REGION Network 17: Sinais Main Line POSTO 80
   // JOB [0]=- ANDON;
   // JOB [1] = EMERGÊNCIA;
   // JOB [2] = AP SUP FREIO;
   // JOB [3] = PY EXCENTRIO;
   // JOB [4] = PY CUBO DISCO
   RUNG wire#powerrail
      Contact( "Get Sinais de Interlock Main line".Station[1]."Sinal do job"[0] )
      I_Contact( "BYPASS_MOD_2" )
      I_Contact( "BYPASS_GERAL" )
      I_Contact( "BYPASS_POSTO_80" )
      Coil( "Signals".ProcessInterlock_APLC_Input[1].ModezoneInterlock_APLC_Input[2].StationInterlock_APLC_Input[3].PositionInterlock_APLC_Input[1].EquipmentInterlock_APLC_Input[1].SignalInterlock_APLC_Input[1] )
   END_RUNG
   RUNG wire#powerrail
      Contact( "Get Sinais de Interlock Main line".Station[1]."Sinal do job"[1] )
      I_Contact( "BYPASS_MOD_2" )
      I_Contact( "BYPASS_GERAL" )
      I_Contact( "BYPASS_POSTO_80" )
      Coil( "Signals".ProcessInterlock_APLC_Input[1].ModezoneInterlock_APLC_Input[2].StationInterlock_APLC_Input[3].PositionInterlock_APLC_Input[1].EquipmentInterlock_APLC_Input[1].SignalInterlock_APLC_Input[2] )
   END_RUNG
   // the same network as SCL:
   "Signals".ProcessInterlock_APLC_Input[1].ModezoneInterlock_APLC_Input[2].StationInterlock_APLC_Input[3].PositionInterlock_APLC_Input[1].EquipmentInterlock_APLC_Input[1].SignalInterlock_APLC_Input[1] := "Get Sinais de Interlock Main line".Station[1]."Sinal do job"[0] AND NOT "BYPASS_MOD_2" AND NOT "BYPASS_GERAL" AND NOT "BYPASS_POSTO_80";
   "Signals".ProcessInterlock_APLC_Input[1].ModezoneInterlock_APLC_Input[2].StationInterlock_APLC_Input[3].PositionInterlock_APLC_Input[1].EquipmentInterlock_APLC_Input[1].SignalInterlock_APLC_Input[2] := "Get Sinais de Interlock Main line".Station[1]."Sinal do job"[1] AND NOT "BYPASS_MOD_2" AND NOT "BYPASS_GERAL" AND NOT "BYPASS_POSTO_80";
END_REGION

REGION Network 18: Sinais Main Line POSTO 90
   // JOB [0] = ANDON;
   // JOB [1] = EMERGÊNCIA;
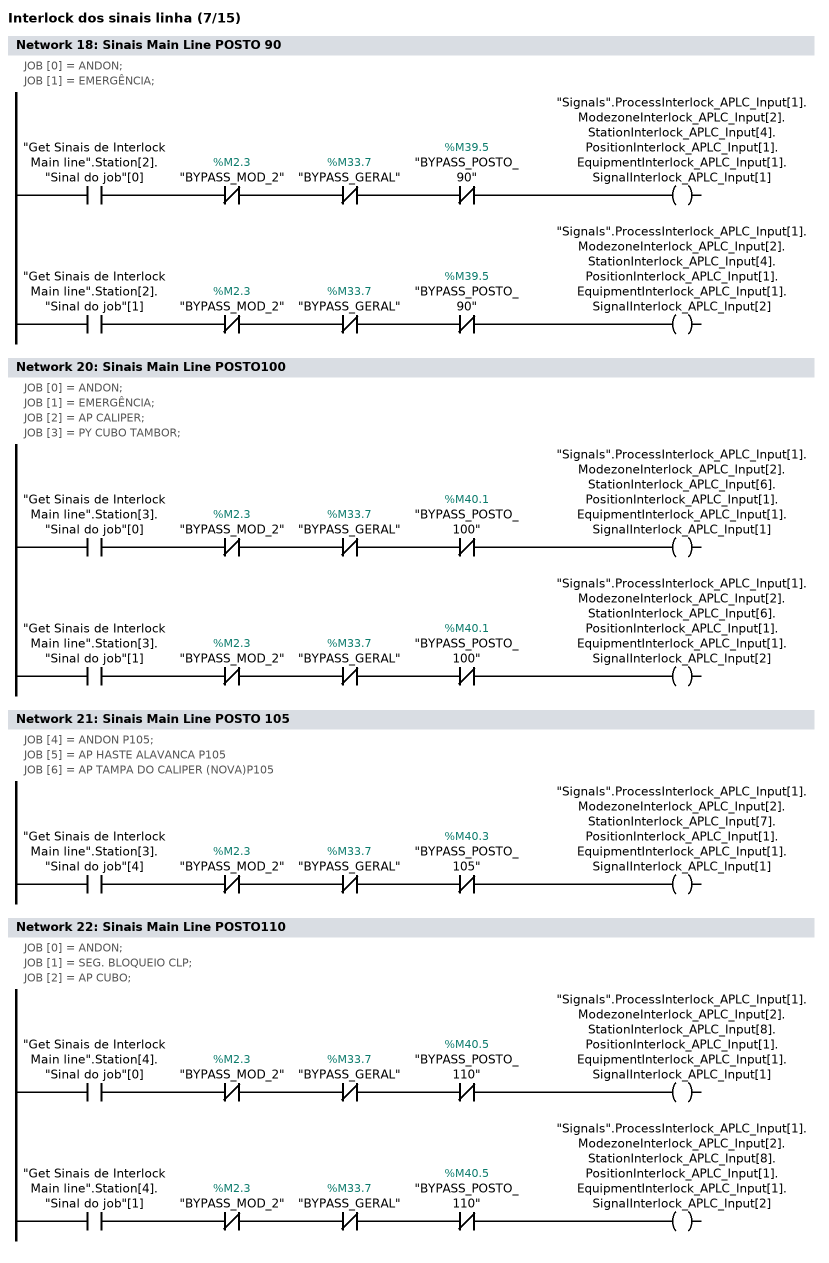
   RUNG wire#powerrail
      Contact( "Get Sinais de Interlock Main line".Station[2]."Sinal do job"[0] )
      I_Contact( "BYPASS_MOD_2" )
      I_Contact( "BYPASS_GERAL" )
      I_Contact( "BYPASS_POSTO_90" )
      Coil( "Signals".ProcessInterlock_APLC_Input[1].ModezoneInterlock_APLC_Input[2].StationInterlock_APLC_Input[4].PositionInterlock_APLC_Input[1].EquipmentInterlock_APLC_Input[1].SignalInterlock_APLC_Input[1] )
   END_RUNG
   RUNG wire#powerrail
      Contact( "Get Sinais de Interlock Main line".Station[2]."Sinal do job"[1] )
      I_Contact( "BYPASS_MOD_2" )
      I_Contact( "BYPASS_GERAL" )
      I_Contact( "BYPASS_POSTO_90" )
      Coil( "Signals".ProcessInterlock_APLC_Input[1].ModezoneInterlock_APLC_Input[2].StationInterlock_APLC_Input[4].PositionInterlock_APLC_Input[1].EquipmentInterlock_APLC_Input[1].SignalInterlock_APLC_Input[2] )
   END_RUNG
   // the same network as SCL:
   "Signals".ProcessInterlock_APLC_Input[1].ModezoneInterlock_APLC_Input[2].StationInterlock_APLC_Input[4].PositionInterlock_APLC_Input[1].EquipmentInterlock_APLC_Input[1].SignalInterlock_APLC_Input[1] := "Get Sinais de Interlock Main line".Station[2]."Sinal do job"[0] AND NOT "BYPASS_MOD_2" AND NOT "BYPASS_GERAL" AND NOT "BYPASS_POSTO_90";
   "Signals".ProcessInterlock_APLC_Input[1].ModezoneInterlock_APLC_Input[2].StationInterlock_APLC_Input[4].PositionInterlock_APLC_Input[1].EquipmentInterlock_APLC_Input[1].SignalInterlock_APLC_Input[2] := "Get Sinais de Interlock Main line".Station[2]."Sinal do job"[1] AND NOT "BYPASS_MOD_2" AND NOT "BYPASS_GERAL" AND NOT "BYPASS_POSTO_90";
END_REGION

REGION Network 19: Sinais Main Line POSTO 95
   // JOB [2] = AP HOLDER. P95
END_REGION

REGION Network 20: Sinais Main Line POSTO100
   // JOB [0] = ANDON;
   // JOB [1] = EMERGÊNCIA;
   // JOB [2] = AP CALIPER;
   // JOB [3] = PY CUBO TAMBOR;
   RUNG wire#powerrail
      Contact( "Get Sinais de Interlock Main line".Station[3]."Sinal do job"[0] )
      I_Contact( "BYPASS_MOD_2" )
      I_Contact( "BYPASS_GERAL" )
      I_Contact( "BYPASS_POSTO_100" )
      Coil( "Signals".ProcessInterlock_APLC_Input[1].ModezoneInterlock_APLC_Input[2].StationInterlock_APLC_Input[6].PositionInterlock_APLC_Input[1].EquipmentInterlock_APLC_Input[1].SignalInterlock_APLC_Input[1] )
   END_RUNG
   RUNG wire#powerrail
      Contact( "Get Sinais de Interlock Main line".Station[3]."Sinal do job"[1] )
      I_Contact( "BYPASS_MOD_2" )
      I_Contact( "BYPASS_GERAL" )
      I_Contact( "BYPASS_POSTO_100" )
      Coil( "Signals".ProcessInterlock_APLC_Input[1].ModezoneInterlock_APLC_Input[2].StationInterlock_APLC_Input[6].PositionInterlock_APLC_Input[1].EquipmentInterlock_APLC_Input[1].SignalInterlock_APLC_Input[2] )
   END_RUNG
   // the same network as SCL:
   "Signals".ProcessInterlock_APLC_Input[1].ModezoneInterlock_APLC_Input[2].StationInterlock_APLC_Input[6].PositionInterlock_APLC_Input[1].EquipmentInterlock_APLC_Input[1].SignalInterlock_APLC_Input[1] := "Get Sinais de Interlock Main line".Station[3]."Sinal do job"[0] AND NOT "BYPASS_MOD_2" AND NOT "BYPASS_GERAL" AND NOT "BYPASS_POSTO_100";
   "Signals".ProcessInterlock_APLC_Input[1].ModezoneInterlock_APLC_Input[2].StationInterlock_APLC_Input[6].PositionInterlock_APLC_Input[1].EquipmentInterlock_APLC_Input[1].SignalInterlock_APLC_Input[2] := "Get Sinais de Interlock Main line".Station[3]."Sinal do job"[1] AND NOT "BYPASS_MOD_2" AND NOT "BYPASS_GERAL" AND NOT "BYPASS_POSTO_100";
END_REGION

REGION Network 21: Sinais Main Line POSTO 105
   // JOB [4] = ANDON P105;
   // JOB [5] = AP HASTE ALAVANCA P105
   // JOB [6] = AP TAMPA DO CALIPER (NOVA)P105
   RUNG wire#powerrail
      Contact( "Get Sinais de Interlock Main line".Station[3]."Sinal do job"[4] )
      I_Contact( "BYPASS_MOD_2" )
      I_Contact( "BYPASS_GERAL" )
      I_Contact( "BYPASS_POSTO_105" )
      Coil( "Signals".ProcessInterlock_APLC_Input[1].ModezoneInterlock_APLC_Input[2].StationInterlock_APLC_Input[7].PositionInterlock_APLC_Input[1].EquipmentInterlock_APLC_Input[1].SignalInterlock_APLC_Input[1] )
   END_RUNG
   // the same network as SCL:
   "Signals".ProcessInterlock_APLC_Input[1].ModezoneInterlock_APLC_Input[2].StationInterlock_APLC_Input[7].PositionInterlock_APLC_Input[1].EquipmentInterlock_APLC_Input[1].SignalInterlock_APLC_Input[1] := "Get Sinais de Interlock Main line".Station[3]."Sinal do job"[4] AND NOT "BYPASS_MOD_2" AND NOT "BYPASS_GERAL" AND NOT "BYPASS_POSTO_105";
END_REGION

REGION Network 22: Sinais Main Line POSTO110
   // JOB [0] = ANDON;
   // JOB [1] = SEG. BLOQUEIO CLP;
   // JOB [2] = AP CUBO;
   RUNG wire#powerrail
      Contact( "Get Sinais de Interlock Main line".Station[4]."Sinal do job"[0] )
      I_Contact( "BYPASS_MOD_2" )
      I_Contact( "BYPASS_GERAL" )
      I_Contact( "BYPASS_POSTO_110" )
      Coil( "Signals".ProcessInterlock_APLC_Input[1].ModezoneInterlock_APLC_Input[2].StationInterlock_APLC_Input[8].PositionInterlock_APLC_Input[1].EquipmentInterlock_APLC_Input[1].SignalInterlock_APLC_Input[1] )
   END_RUNG
   RUNG wire#powerrail
      Contact( "Get Sinais de Interlock Main line".Station[4]."Sinal do job"[1] )
      I_Contact( "BYPASS_MOD_2" )
      I_Contact( "BYPASS_GERAL" )
      I_Contact( "BYPASS_POSTO_110" )
      Coil( "Signals".ProcessInterlock_APLC_Input[1].ModezoneInterlock_APLC_Input[2].StationInterlock_APLC_Input[8].PositionInterlock_APLC_Input[1].EquipmentInterlock_APLC_Input[1].SignalInterlock_APLC_Input[2] )
   END_RUNG
   // the same network as SCL:
   "Signals".ProcessInterlock_APLC_Input[1].ModezoneInterlock_APLC_Input[2].StationInterlock_APLC_Input[8].PositionInterlock_APLC_Input[1].EquipmentInterlock_APLC_Input[1].SignalInterlock_APLC_Input[1] := "Get Sinais de Interlock Main line".Station[4]."Sinal do job"[0] AND NOT "BYPASS_MOD_2" AND NOT "BYPASS_GERAL" AND NOT "BYPASS_POSTO_110";
   "Signals".ProcessInterlock_APLC_Input[1].ModezoneInterlock_APLC_Input[2].StationInterlock_APLC_Input[8].PositionInterlock_APLC_Input[1].EquipmentInterlock_APLC_Input[1].SignalInterlock_APLC_Input[2] := "Get Sinais de Interlock Main line".Station[4]."Sinal do job"[1] AND NOT "BYPASS_MOD_2" AND NOT "BYPASS_GERAL" AND NOT "BYPASS_POSTO_110";
END_REGION

REGION Network 23: Sinais Main Line POSTO 115
   // JOB [3] = ANDON P115;
   // JOB [4] = CRAVADOR.
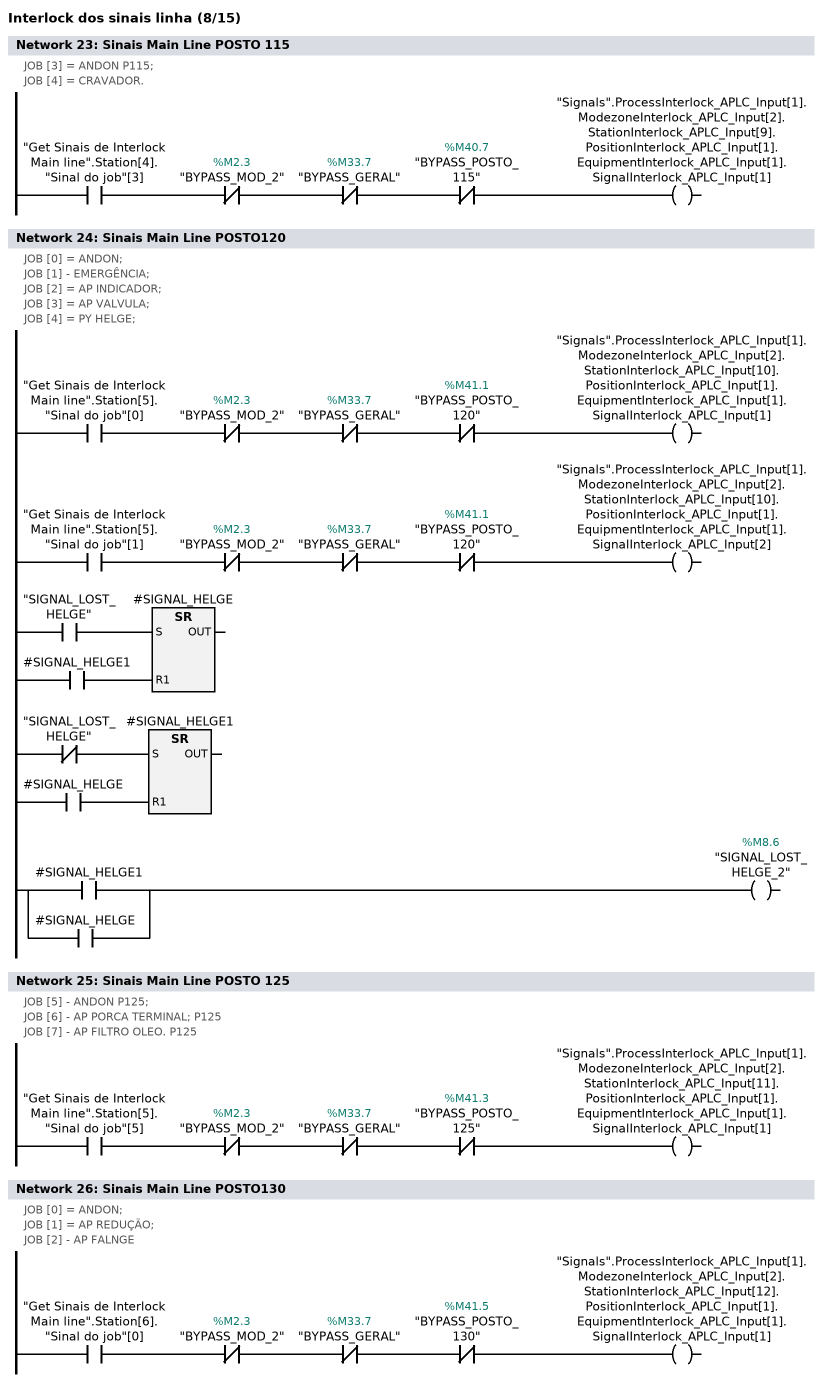
   RUNG wire#powerrail
      Contact( "Get Sinais de Interlock Main line".Station[4]."Sinal do job"[3] )
      I_Contact( "BYPASS_MOD_2" )
      I_Contact( "BYPASS_GERAL" )
      I_Contact( "BYPASS_POSTO_115" )
      Coil( "Signals".ProcessInterlock_APLC_Input[1].ModezoneInterlock_APLC_Input[2].StationInterlock_APLC_Input[9].PositionInterlock_APLC_Input[1].EquipmentInterlock_APLC_Input[1].SignalInterlock_APLC_Input[1] )
   END_RUNG
   // the same network as SCL:
   "Signals".ProcessInterlock_APLC_Input[1].ModezoneInterlock_APLC_Input[2].StationInterlock_APLC_Input[9].PositionInterlock_APLC_Input[1].EquipmentInterlock_APLC_Input[1].SignalInterlock_APLC_Input[1] := "Get Sinais de Interlock Main line".Station[4]."Sinal do job"[3] AND NOT "BYPASS_MOD_2" AND NOT "BYPASS_GERAL" AND NOT "BYPASS_POSTO_115";
END_REGION

REGION Network 24: Sinais Main Line POSTO120
   // JOB [0] = ANDON;
   // JOB [1] - EMERGÊNCIA;
   // JOB [2] = AP INDICADOR;
   // JOB [3] = AP VALVULA;
   // JOB [4] = PY HELGE;
   RUNG wire#powerrail
      Contact( "Get Sinais de Interlock Main line".Station[5]."Sinal do job"[0] )
      I_Contact( "BYPASS_MOD_2" )
      I_Contact( "BYPASS_GERAL" )
      I_Contact( "BYPASS_POSTO_120" )
      Coil( "Signals".ProcessInterlock_APLC_Input[1].ModezoneInterlock_APLC_Input[2].StationInterlock_APLC_Input[10].PositionInterlock_APLC_Input[1].EquipmentInterlock_APLC_Input[1].SignalInterlock_APLC_Input[1] )
   END_RUNG
   RUNG wire#powerrail
      Contact( "Get Sinais de Interlock Main line".Station[5]."Sinal do job"[1] )
      I_Contact( "BYPASS_MOD_2" )
      I_Contact( "BYPASS_GERAL" )
      I_Contact( "BYPASS_POSTO_120" )
      Coil( "Signals".ProcessInterlock_APLC_Input[1].ModezoneInterlock_APLC_Input[2].StationInterlock_APLC_Input[10].PositionInterlock_APLC_Input[1].EquipmentInterlock_APLC_Input[1].SignalInterlock_APLC_Input[2] )
   END_RUNG
   RUNG wire#powerrail
      Contact( "SIGNAL_LOST_HELGE" )
      S_SR(operand := #SIGNAL_HELGE, r1 := wire#w1)
   END_RUNG
   RUNG wire#powerrail
      Contact( #SIGNAL_HELGE1 )
   END_RUNG wire#w1
   RUNG wire#powerrail
      I_Contact( "SIGNAL_LOST_HELGE" )
      S_SR(operand := #SIGNAL_HELGE1, r1 := wire#w2)
   END_RUNG
   RUNG wire#powerrail
      Contact( #SIGNAL_HELGE )
   END_RUNG wire#w2
   RUNG wire#powerrail
      Contact( #SIGNAL_HELGE1 )
      wire#w3
      Coil( "SIGNAL_LOST_HELGE_2" )
   END_RUNG
   RUNG wire#powerrail
      Contact( #SIGNAL_HELGE )
   END_RUNG wire#w3
   // the same network as SCL:
   "Signals".ProcessInterlock_APLC_Input[1].ModezoneInterlock_APLC_Input[2].StationInterlock_APLC_Input[10].PositionInterlock_APLC_Input[1].EquipmentInterlock_APLC_Input[1].SignalInterlock_APLC_Input[1] := "Get Sinais de Interlock Main line".Station[5]."Sinal do job"[0] AND NOT "BYPASS_MOD_2" AND NOT "BYPASS_GERAL" AND NOT "BYPASS_POSTO_120";
   "Signals".ProcessInterlock_APLC_Input[1].ModezoneInterlock_APLC_Input[2].StationInterlock_APLC_Input[10].PositionInterlock_APLC_Input[1].EquipmentInterlock_APLC_Input[1].SignalInterlock_APLC_Input[2] := "Get Sinais de Interlock Main line".Station[5]."Sinal do job"[1] AND NOT "BYPASS_MOD_2" AND NOT "BYPASS_GERAL" AND NOT "BYPASS_POSTO_120";
   IF "SIGNAL_LOST_HELGE" THEN
       #SIGNAL_HELGE := TRUE;   // SR flip-flop
   END_IF;
   IF #SIGNAL_HELGE1 THEN #SIGNAL_HELGE := FALSE; END_IF;
   IF NOT "SIGNAL_LOST_HELGE" THEN
       #SIGNAL_HELGE1 := TRUE;   // SR flip-flop
   END_IF;
   IF #SIGNAL_HELGE THEN #SIGNAL_HELGE1 := FALSE; END_IF;
   "SIGNAL_LOST_HELGE_2" := #SIGNAL_HELGE1 OR #SIGNAL_HELGE;
END_REGION

REGION Network 25: Sinais Main Line POSTO 125
   // JOB [5] - ANDON P125;
   // JOB [6] - AP PORCA TERMINAL; P125
   // JOB [7] - AP FILTRO OLEO. P125
   RUNG wire#powerrail
      Contact( "Get Sinais de Interlock Main line".Station[5]."Sinal do job"[5] )
      I_Contact( "BYPASS_MOD_2" )
      I_Contact( "BYPASS_GERAL" )
      I_Contact( "BYPASS_POSTO_125" )
      Coil( "Signals".ProcessInterlock_APLC_Input[1].ModezoneInterlock_APLC_Input[2].StationInterlock_APLC_Input[11].PositionInterlock_APLC_Input[1].EquipmentInterlock_APLC_Input[1].SignalInterlock_APLC_Input[1] )
   END_RUNG
   // the same network as SCL:
   "Signals".ProcessInterlock_APLC_Input[1].ModezoneInterlock_APLC_Input[2].StationInterlock_APLC_Input[11].PositionInterlock_APLC_Input[1].EquipmentInterlock_APLC_Input[1].SignalInterlock_APLC_Input[1] := "Get Sinais de Interlock Main line".Station[5]."Sinal do job"[5] AND NOT "BYPASS_MOD_2" AND NOT "BYPASS_GERAL" AND NOT "BYPASS_POSTO_125";
END_REGION

REGION Network 26: Sinais Main Line POSTO130
   // JOB [0] = ANDON;
   // JOB [1] = AP REDUÇÃO;
   // JOB [2] - AP FALNGE
   RUNG wire#powerrail
      Contact( "Get Sinais de Interlock Main line".Station[6]."Sinal do job"[0] )
      I_Contact( "BYPASS_MOD_2" )
      I_Contact( "BYPASS_GERAL" )
      I_Contact( "BYPASS_POSTO_130" )
      Coil( "Signals".ProcessInterlock_APLC_Input[1].ModezoneInterlock_APLC_Input[2].StationInterlock_APLC_Input[12].PositionInterlock_APLC_Input[1].EquipmentInterlock_APLC_Input[1].SignalInterlock_APLC_Input[1] )
   END_RUNG
   // the same network as SCL:
   "Signals".ProcessInterlock_APLC_Input[1].ModezoneInterlock_APLC_Input[2].StationInterlock_APLC_Input[12].PositionInterlock_APLC_Input[1].EquipmentInterlock_APLC_Input[1].SignalInterlock_APLC_Input[1] := "Get Sinais de Interlock Main line".Station[6]."Sinal do job"[0] AND NOT "BYPASS_MOD_2" AND NOT "BYPASS_GERAL" AND NOT "BYPASS_POSTO_130";
END_REGION

REGION Network 27: Sinais Main Line POSTO140
   // JOB [0] = ANDON;
   // JOB [1] = EMERGÊNCIA;
   // JOB [2] = ESTANQUEIDADE CILINDRO;
   // JOB [3] = ESTANQUEIDADE CARCAÇA.
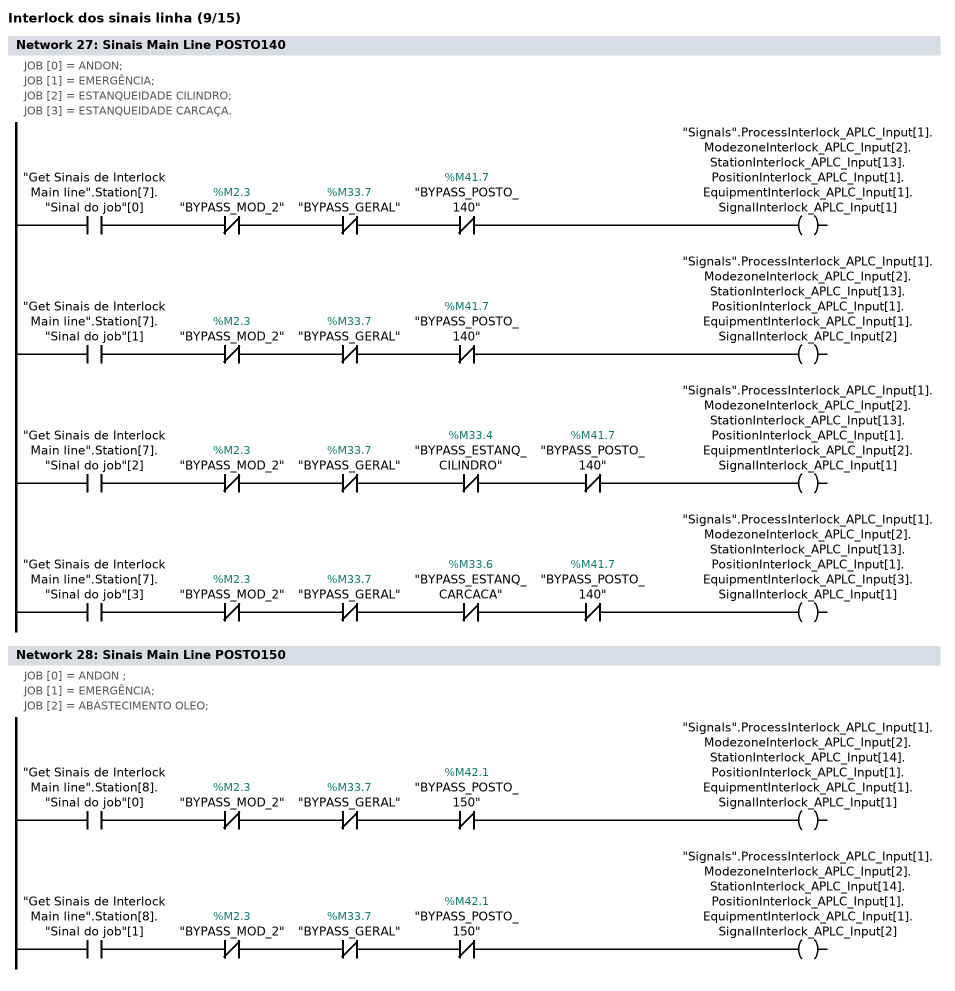
   RUNG wire#powerrail
      Contact( "Get Sinais de Interlock Main line".Station[7]."Sinal do job"[0] )
      I_Contact( "BYPASS_MOD_2" )
      I_Contact( "BYPASS_GERAL" )
      I_Contact( "BYPASS_POSTO_140" )
      Coil( "Signals".ProcessInterlock_APLC_Input[1].ModezoneInterlock_APLC_Input[2].StationInterlock_APLC_Input[13].PositionInterlock_APLC_Input[1].EquipmentInterlock_APLC_Input[1].SignalInterlock_APLC_Input[1] )
   END_RUNG
   RUNG wire#powerrail
      Contact( "Get Sinais de Interlock Main line".Station[7]."Sinal do job"[1] )
      I_Contact( "BYPASS_MOD_2" )
      I_Contact( "BYPASS_GERAL" )
      I_Contact( "BYPASS_POSTO_140" )
      Coil( "Signals".ProcessInterlock_APLC_Input[1].ModezoneInterlock_APLC_Input[2].StationInterlock_APLC_Input[13].PositionInterlock_APLC_Input[1].EquipmentInterlock_APLC_Input[1].SignalInterlock_APLC_Input[2] )
   END_RUNG
   RUNG wire#powerrail
      Contact( "Get Sinais de Interlock Main line".Station[7]."Sinal do job"[2] )
      I_Contact( "BYPASS_MOD_2" )
      I_Contact( "BYPASS_GERAL" )
      I_Contact( "BYPASS_ESTANQ_CILINDRO" )
      I_Contact( "BYPASS_POSTO_140" )
      Coil( "Signals".ProcessInterlock_APLC_Input[1].ModezoneInterlock_APLC_Input[2].StationInterlock_APLC_Input[13].PositionInterlock_APLC_Input[1].EquipmentInterlock_APLC_Input[2].SignalInterlock_APLC_Input[1] )
   END_RUNG
   RUNG wire#powerrail
      Contact( "Get Sinais de Interlock Main line".Station[7]."Sinal do job"[3] )
      I_Contact( "BYPASS_MOD_2" )
      I_Contact( "BYPASS_GERAL" )
      I_Contact( "BYPASS_ESTANQ_CARCACA" )
      I_Contact( "BYPASS_POSTO_140" )
      Coil( "Signals".ProcessInterlock_APLC_Input[1].ModezoneInterlock_APLC_Input[2].StationInterlock_APLC_Input[13].PositionInterlock_APLC_Input[1].EquipmentInterlock_APLC_Input[3].SignalInterlock_APLC_Input[1] )
   END_RUNG
   // the same network as SCL:
   "Signals".ProcessInterlock_APLC_Input[1].ModezoneInterlock_APLC_Input[2].StationInterlock_APLC_Input[13].PositionInterlock_APLC_Input[1].EquipmentInterlock_APLC_Input[1].SignalInterlock_APLC_Input[1] := "Get Sinais de Interlock Main line".Station[7]."Sinal do job"[0] AND NOT "BYPASS_MOD_2" AND NOT "BYPASS_GERAL" AND NOT "BYPASS_POSTO_140";
   "Signals".ProcessInterlock_APLC_Input[1].ModezoneInterlock_APLC_Input[2].StationInterlock_APLC_Input[13].PositionInterlock_APLC_Input[1].EquipmentInterlock_APLC_Input[1].SignalInterlock_APLC_Input[2] := "Get Sinais de Interlock Main line".Station[7]."Sinal do job"[1] AND NOT "BYPASS_MOD_2" AND NOT "BYPASS_GERAL" AND NOT "BYPASS_POSTO_140";
   "Signals".ProcessInterlock_APLC_Input[1].ModezoneInterlock_APLC_Input[2].StationInterlock_APLC_Input[13].PositionInterlock_APLC_Input[1].EquipmentInterlock_APLC_Input[2].SignalInterlock_APLC_Input[1] := "Get Sinais de Interlock Main line".Station[7]."Sinal do job"[2] AND NOT "BYPASS_MOD_2" AND NOT "BYPASS_GERAL" AND NOT "BYPASS_ESTANQ_CILINDRO" AND NOT "BYPASS_POSTO_140";
   "Signals".ProcessInterlock_APLC_Input[1].ModezoneInterlock_APLC_Input[2].StationInterlock_APLC_Input[13].PositionInterlock_APLC_Input[1].EquipmentInterlock_APLC_Input[3].SignalInterlock_APLC_Input[1] := "Get Sinais de Interlock Main line".Station[7]."Sinal do job"[3] AND NOT "BYPASS_MOD_2" AND NOT "BYPASS_GERAL" AND NOT "BYPASS_ESTANQ_CARCACA" AND NOT "BYPASS_POSTO_140";
END_REGION

REGION Network 28: Sinais Main Line POSTO150
   // JOB [0] = ANDON ;
   // JOB [1] = EMERGÊNCIA;
   // JOB [2] = ABASTECIMENTO OLEO;
   RUNG wire#powerrail
      Contact( "Get Sinais de Interlock Main line".Station[8]."Sinal do job"[0] )
      I_Contact( "BYPASS_MOD_2" )
      I_Contact( "BYPASS_GERAL" )
      I_Contact( "BYPASS_POSTO_150" )
      Coil( "Signals".ProcessInterlock_APLC_Input[1].ModezoneInterlock_APLC_Input[2].StationInterlock_APLC_Input[14].PositionInterlock_APLC_Input[1].EquipmentInterlock_APLC_Input[1].SignalInterlock_APLC_Input[1] )
   END_RUNG
   RUNG wire#powerrail
      Contact( "Get Sinais de Interlock Main line".Station[8]."Sinal do job"[1] )
      I_Contact( "BYPASS_MOD_2" )
      I_Contact( "BYPASS_GERAL" )
      I_Contact( "BYPASS_POSTO_150" )
      Coil( "Signals".ProcessInterlock_APLC_Input[1].ModezoneInterlock_APLC_Input[2].StationInterlock_APLC_Input[14].PositionInterlock_APLC_Input[1].EquipmentInterlock_APLC_Input[1].SignalInterlock_APLC_Input[2] )
   END_RUNG
   // the same network as SCL:
   "Signals".ProcessInterlock_APLC_Input[1].ModezoneInterlock_APLC_Input[2].StationInterlock_APLC_Input[14].PositionInterlock_APLC_Input[1].EquipmentInterlock_APLC_Input[1].SignalInterlock_APLC_Input[1] := "Get Sinais de Interlock Main line".Station[8]."Sinal do job"[0] AND NOT "BYPASS_MOD_2" AND NOT "BYPASS_GERAL" AND NOT "BYPASS_POSTO_150";
   "Signals".ProcessInterlock_APLC_Input[1].ModezoneInterlock_APLC_Input[2].StationInterlock_APLC_Input[14].PositionInterlock_APLC_Input[1].EquipmentInterlock_APLC_Input[1].SignalInterlock_APLC_Input[2] := "Get Sinais de Interlock Main line".Station[8]."Sinal do job"[1] AND NOT "BYPASS_MOD_2" AND NOT "BYPASS_GERAL" AND NOT "BYPASS_POSTO_150";
END_REGION

REGION Network 29: Sinais Main Line Q.G
   // JOB [0] = ANDON;
   // JOB [1] = EMERGÊNCIA;
   // JOB [2] - EIXO PENDURADO;
   // JOB [3] - GAP PRESENTE CAB;
   // JOB [4] - GAP PRESENTE TAKT 
   // STATION 10 JOB [0] = TRANSPORTADOR EM MANUAL
   // GAP + EIXO PENDURADO
   // MODEZONE 1 PARADO (FALCARE)
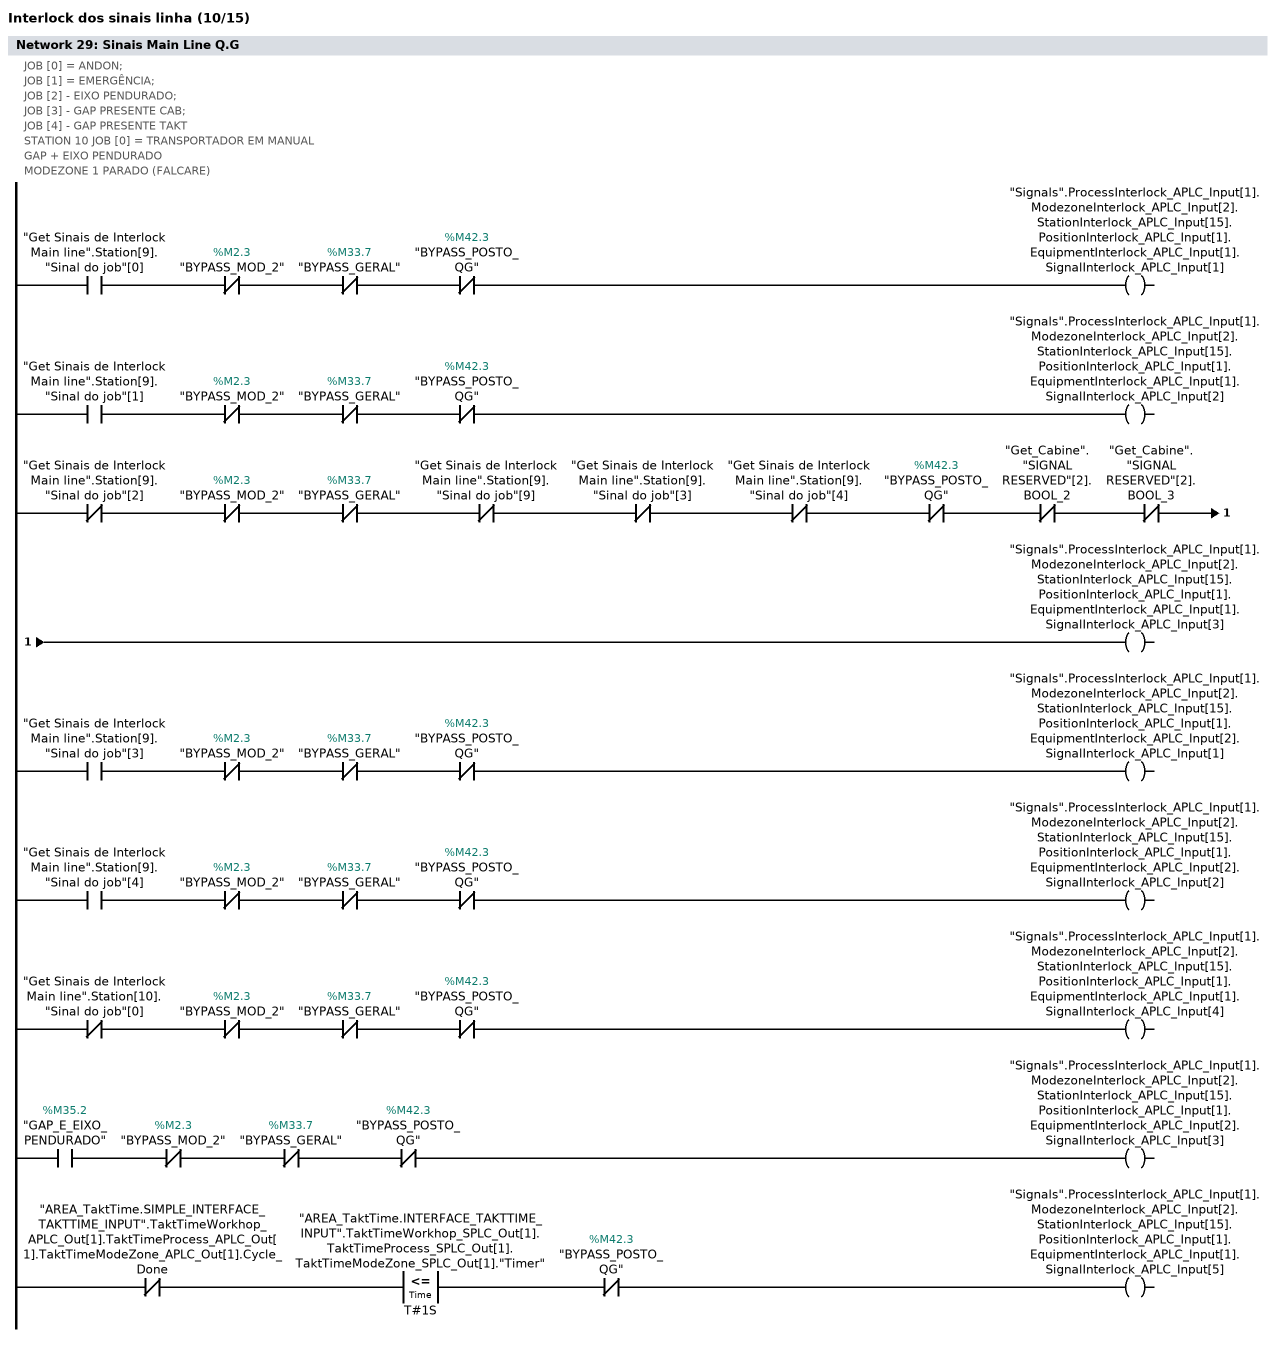
   RUNG wire#powerrail
      Contact( "Get Sinais de Interlock Main line".Station[9]."Sinal do job"[0] )
      I_Contact( "BYPASS_MOD_2" )
      I_Contact( "BYPASS_GERAL" )
      I_Contact( "BYPASS_POSTO_QG" )
      Coil( "Signals".ProcessInterlock_APLC_Input[1].ModezoneInterlock_APLC_Input[2].StationInterlock_APLC_Input[15].PositionInterlock_APLC_Input[1].EquipmentInterlock_APLC_Input[1].SignalInterlock_APLC_Input[1] )
   END_RUNG
   RUNG wire#powerrail
      Contact( "Get Sinais de Interlock Main line".Station[9]."Sinal do job"[1] )
      I_Contact( "BYPASS_MOD_2" )
      I_Contact( "BYPASS_GERAL" )
      I_Contact( "BYPASS_POSTO_QG" )
      Coil( "Signals".ProcessInterlock_APLC_Input[1].ModezoneInterlock_APLC_Input[2].StationInterlock_APLC_Input[15].PositionInterlock_APLC_Input[1].EquipmentInterlock_APLC_Input[1].SignalInterlock_APLC_Input[2] )
   END_RUNG
   RUNG wire#powerrail
      I_Contact( "Get Sinais de Interlock Main line".Station[9]."Sinal do job"[2] )
      I_Contact( "BYPASS_MOD_2" )
      I_Contact( "BYPASS_GERAL" )
      I_Contact( "Get Sinais de Interlock Main line".Station[9]."Sinal do job"[9] )
      I_Contact( "Get Sinais de Interlock Main line".Station[9]."Sinal do job"[3] )
      I_Contact( "Get Sinais de Interlock Main line".Station[9]."Sinal do job"[4] )
      I_Contact( "BYPASS_POSTO_QG" )
      I_Contact( "Get_Cabine"."SIGNAL RESERVED"[2].BOOL_2 )
      I_Contact( "Get_Cabine"."SIGNAL RESERVED"[2].BOOL_3 )
      Coil( "Signals".ProcessInterlock_APLC_Input[1].ModezoneInterlock_APLC_Input[2].StationInterlock_APLC_Input[15].PositionInterlock_APLC_Input[1].EquipmentInterlock_APLC_Input[1].SignalInterlock_APLC_Input[3] )
   END_RUNG
   RUNG wire#powerrail
      Contact( "Get Sinais de Interlock Main line".Station[9]."Sinal do job"[3] )
      I_Contact( "BYPASS_MOD_2" )
      I_Contact( "BYPASS_GERAL" )
      I_Contact( "BYPASS_POSTO_QG" )
      Coil( "Signals".ProcessInterlock_APLC_Input[1].ModezoneInterlock_APLC_Input[2].StationInterlock_APLC_Input[15].PositionInterlock_APLC_Input[1].EquipmentInterlock_APLC_Input[2].SignalInterlock_APLC_Input[1] )
   END_RUNG
   RUNG wire#powerrail
      Contact( "Get Sinais de Interlock Main line".Station[9]."Sinal do job"[4] )
      I_Contact( "BYPASS_MOD_2" )
      I_Contact( "BYPASS_GERAL" )
      I_Contact( "BYPASS_POSTO_QG" )
      Coil( "Signals".ProcessInterlock_APLC_Input[1].ModezoneInterlock_APLC_Input[2].StationInterlock_APLC_Input[15].PositionInterlock_APLC_Input[1].EquipmentInterlock_APLC_Input[2].SignalInterlock_APLC_Input[2] )
   END_RUNG
   RUNG wire#powerrail
      I_Contact( "Get Sinais de Interlock Main line".Station[10]."Sinal do job"[0] )
      I_Contact( "BYPASS_MOD_2" )
      I_Contact( "BYPASS_GERAL" )
      I_Contact( "BYPASS_POSTO_QG" )
      Coil( "Signals".ProcessInterlock_APLC_Input[1].ModezoneInterlock_APLC_Input[2].StationInterlock_APLC_Input[15].PositionInterlock_APLC_Input[1].EquipmentInterlock_APLC_Input[1].SignalInterlock_APLC_Input[4] )
   END_RUNG
   RUNG wire#powerrail
      Contact( "GAP_E_EIXO_PENDURADO" )
      I_Contact( "BYPASS_MOD_2" )
      I_Contact( "BYPASS_GERAL" )
      I_Contact( "BYPASS_POSTO_QG" )
      Coil( "Signals".ProcessInterlock_APLC_Input[1].ModezoneInterlock_APLC_Input[2].StationInterlock_APLC_Input[15].PositionInterlock_APLC_Input[1].EquipmentInterlock_APLC_Input[2].SignalInterlock_APLC_Input[3] )
   END_RUNG
   RUNG wire#powerrail
      I_Contact( "AREA_TaktTime.SIMPLE_INTERFACE_TAKTTIME_INPUT".TaktTimeWorkhop_APLC_Out[1].TaktTimeProcess_APLC_Out[1].TaktTimeModeZone_APLC_Out[1].Cycle_Done )
      { S7_Templates := "SrcType := Time" } LE_Contact(in1 := "AREA_TaktTime.INTERFACE_TAKTTIME_INPUT".TaktTimeWorkhop_SPLC_Out[1].TaktTimeProcess_SPLC_Out[1].TaktTimeModeZone_SPLC_Out[1]."Timer", in2 := T#1S)
      I_Contact( "BYPASS_POSTO_QG" )
      Coil( "Signals".ProcessInterlock_APLC_Input[1].ModezoneInterlock_APLC_Input[2].StationInterlock_APLC_Input[15].PositionInterlock_APLC_Input[1].EquipmentInterlock_APLC_Input[1].SignalInterlock_APLC_Input[5] )
   END_RUNG
   // the same network as SCL:
   "Signals".ProcessInterlock_APLC_Input[1].ModezoneInterlock_APLC_Input[2].StationInterlock_APLC_Input[15].PositionInterlock_APLC_Input[1].EquipmentInterlock_APLC_Input[1].SignalInterlock_APLC_Input[1] := "Get Sinais de Interlock Main line".Station[9]."Sinal do job"[0] AND NOT "BYPASS_MOD_2" AND NOT "BYPASS_GERAL" AND NOT "BYPASS_POSTO_QG";
   "Signals".ProcessInterlock_APLC_Input[1].ModezoneInterlock_APLC_Input[2].StationInterlock_APLC_Input[15].PositionInterlock_APLC_Input[1].EquipmentInterlock_APLC_Input[1].SignalInterlock_APLC_Input[2] := "Get Sinais de Interlock Main line".Station[9]."Sinal do job"[1] AND NOT "BYPASS_MOD_2" AND NOT "BYPASS_GERAL" AND NOT "BYPASS_POSTO_QG";
   "Signals".ProcessInterlock_APLC_Input[1].ModezoneInterlock_APLC_Input[2].StationInterlock_APLC_Input[15].PositionInterlock_APLC_Input[1].EquipmentInterlock_APLC_Input[1].SignalInterlock_APLC_Input[3] := NOT "Get Sinais de Interlock Main line".Station[9]."Sinal do job"[2] AND NOT "BYPASS_MOD_2" AND NOT "BYPASS_GERAL" AND NOT "Get Sinais de Interlock Main line".Station[9]."Sinal do job"[9] AND NOT "Get Sinais de Interlock Main line".Station[9]."Sinal do job"[3] AND NOT "Get Sinais de Interlock Main line".Station[9]."Sinal do job"[4] AND NOT "BYPASS_POSTO_QG" AND NOT "Get_Cabine"."SIGNAL RESERVED"[2].BOOL_2 AND NOT "Get_Cabine"."SIGNAL RESERVED"[2].BOOL_3;
   "Signals".ProcessInterlock_APLC_Input[1].ModezoneInterlock_APLC_Input[2].StationInterlock_APLC_Input[15].PositionInterlock_APLC_Input[1].EquipmentInterlock_APLC_Input[2].SignalInterlock_APLC_Input[1] := "Get Sinais de Interlock Main line".Station[9]."Sinal do job"[3] AND NOT "BYPASS_MOD_2" AND NOT "BYPASS_GERAL" AND NOT "BYPASS_POSTO_QG";
   "Signals".ProcessInterlock_APLC_Input[1].ModezoneInterlock_APLC_Input[2].StationInterlock_APLC_Input[15].PositionInterlock_APLC_Input[1].EquipmentInterlock_APLC_Input[2].SignalInterlock_APLC_Input[2] := "Get Sinais de Interlock Main line".Station[9]."Sinal do job"[4] AND NOT "BYPASS_MOD_2" AND NOT "BYPASS_GERAL" AND NOT "BYPASS_POSTO_QG";
   "Signals".ProcessInterlock_APLC_Input[1].ModezoneInterlock_APLC_Input[2].StationInterlock_APLC_Input[15].PositionInterlock_APLC_Input[1].EquipmentInterlock_APLC_Input[1].SignalInterlock_APLC_Input[4] := NOT "Get Sinais de Interlock Main line".Station[10]."Sinal do job"[0] AND NOT "BYPASS_MOD_2" AND NOT "BYPASS_GERAL" AND NOT "BYPASS_POSTO_QG";
   "Signals".ProcessInterlock_APLC_Input[1].ModezoneInterlock_APLC_Input[2].StationInterlock_APLC_Input[15].PositionInterlock_APLC_Input[1].EquipmentInterlock_APLC_Input[2].SignalInterlock_APLC_Input[3] := "GAP_E_EIXO_PENDURADO" AND NOT "BYPASS_MOD_2" AND NOT "BYPASS_GERAL" AND NOT "BYPASS_POSTO_QG";
   "Signals".ProcessInterlock_APLC_Input[1].ModezoneInterlock_APLC_Input[2].StationInterlock_APLC_Input[15].PositionInterlock_APLC_Input[1].EquipmentInterlock_APLC_Input[1].SignalInterlock_APLC_Input[5] := NOT "AREA_TaktTime.SIMPLE_INTERFACE_TAKTTIME_INPUT".TaktTimeWorkhop_APLC_Out[1].TaktTimeProcess_APLC_Out[1].TaktTimeModeZone_APLC_Out[1].Cycle_Done AND ("AREA_TaktTime.INTERFACE_TAKTTIME_INPUT".TaktTimeWorkhop_SPLC_Out[1].TaktTimeProcess_SPLC_Out[1].TaktTimeModeZone_SPLC_Out[1]."Timer" <= T#1S) AND NOT "BYPASS_POSTO_QG";
END_REGION

REGION Network 30: CABINE DEPINTURA
   // ANDON
   // EMERGÊNCIA
   // PORTAS DA CABINE 
   // SINAL OK DO ROBO (SINAL INFORMANDO QUE A PINTURA FOI CONCLUIDA)
   // TALHA FORA DE POSIÇÃO
   // CABINE NOK (INFORMA QUE TEM ALGUMA FALHA NA CABINE)
   // CONFIRMAÇÃO DE RECEITA
   // TAKT LOCAL
   // SIGNAL RESERVED [1] [BOOL ] = ANDON EXPEDIÇÃO
   // SIGNAL RESERVED [1] [BOOL 1] = ESVAZIAMENTO DE LINHA CABINE
   // SIGNAL RESERVED [1] [BOOL 2] = PLATAFORMA
   // SIGNAL RESERVED [1] [BOOL 3] = ANDON CARGA PLATAFORMA
   // SIGNAL RESERVED [2] [BOOL ] = CABINE GIRANDO
   // SIGNAL RESERVED [2] [BOOL 1 ] = SENSOR DE COLISÃO EXPEDIÇÃO
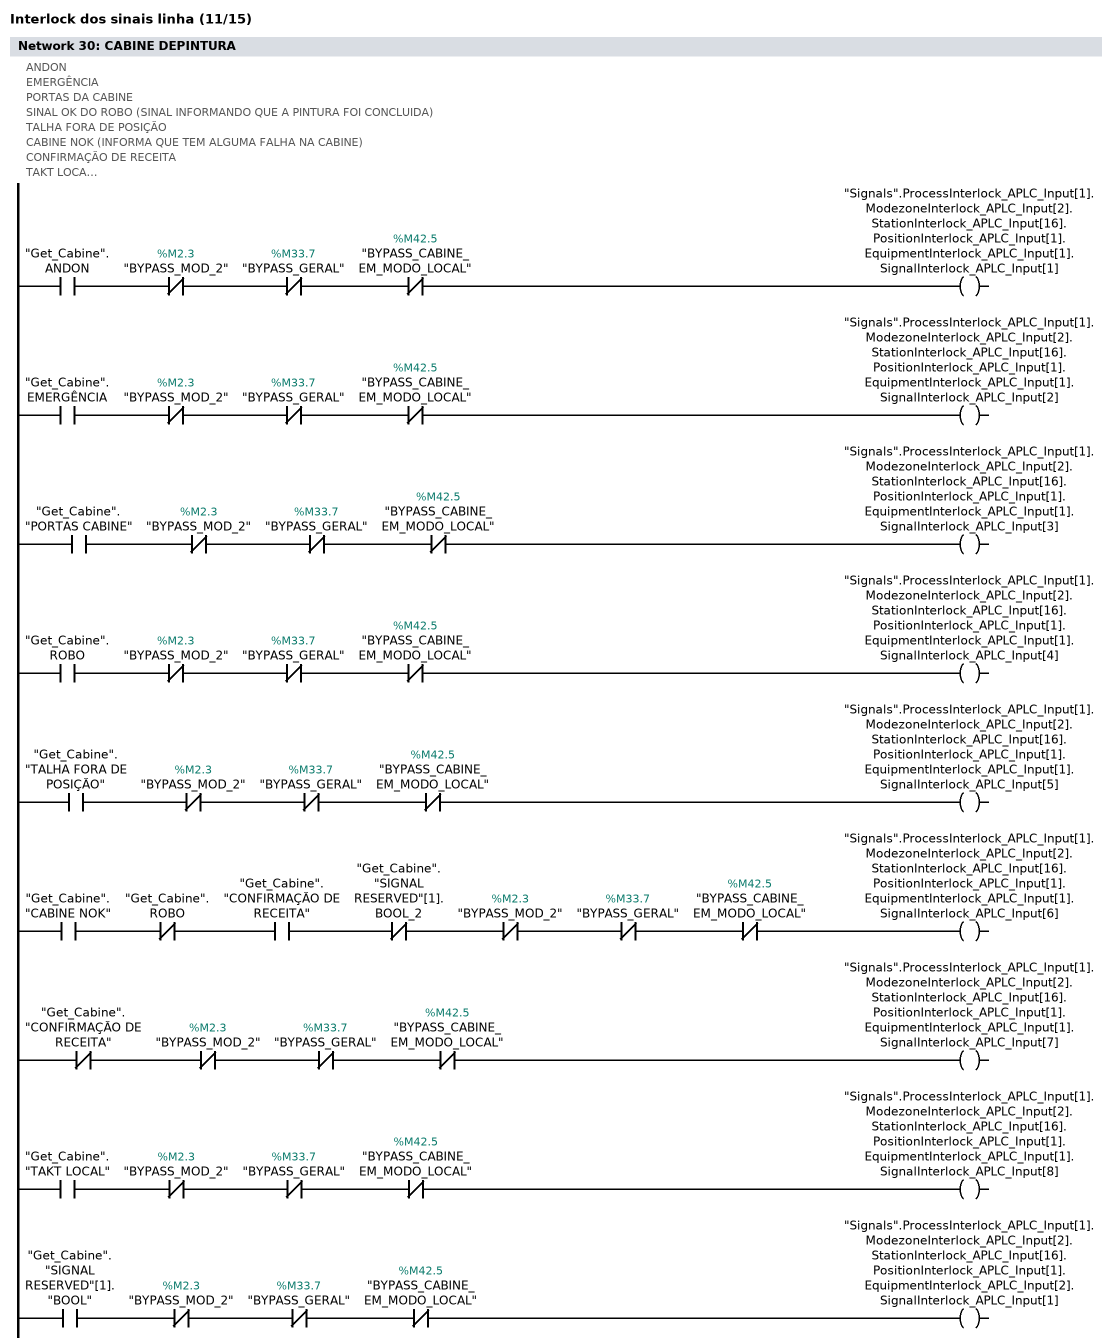
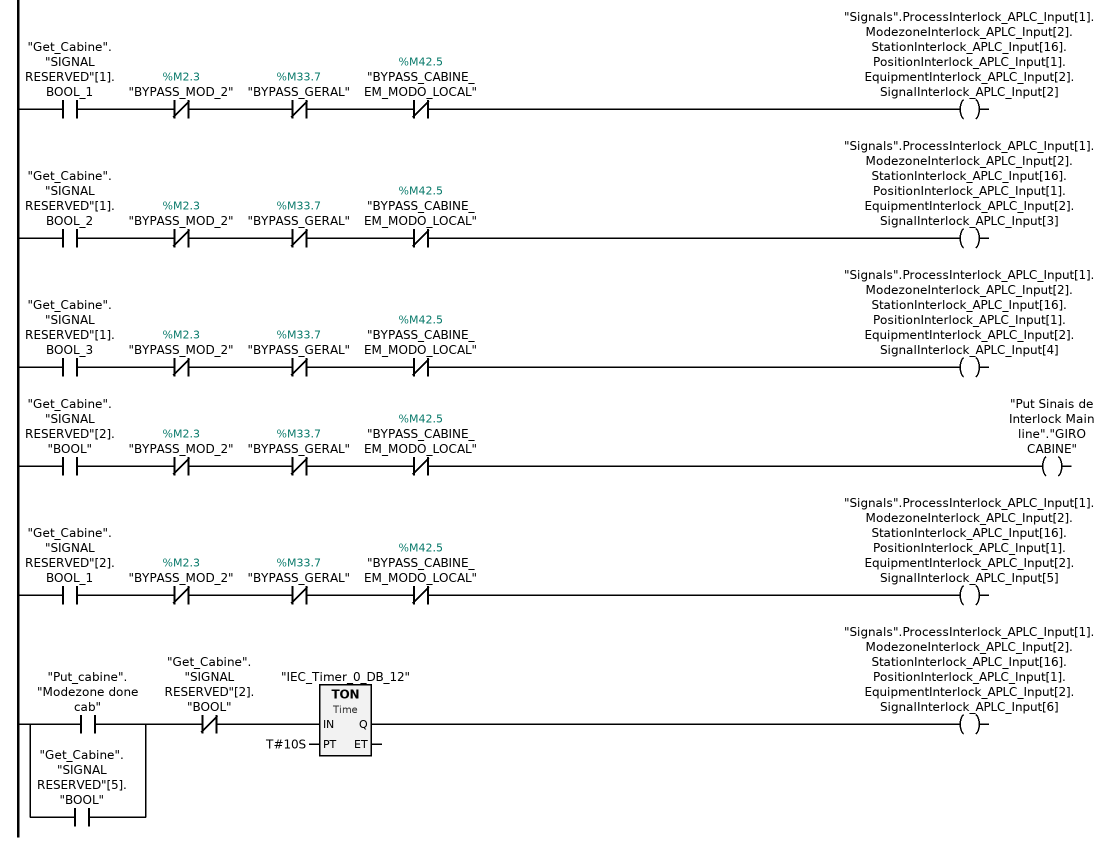
   RUNG wire#powerrail
      Contact( "Get_Cabine".ANDON )
      I_Contact( "BYPASS_MOD_2" )
      I_Contact( "BYPASS_GERAL" )
      I_Contact( "BYPASS_CABINE_EM_MODO_LOCAL" )
      Coil( "Signals".ProcessInterlock_APLC_Input[1].ModezoneInterlock_APLC_Input[2].StationInterlock_APLC_Input[16].PositionInterlock_APLC_Input[1].EquipmentInterlock_APLC_Input[1].SignalInterlock_APLC_Input[1] )
   END_RUNG
   RUNG wire#powerrail
      Contact( "Get_Cabine".EMERGÊNCIA )
      I_Contact( "BYPASS_MOD_2" )
      I_Contact( "BYPASS_GERAL" )
      I_Contact( "BYPASS_CABINE_EM_MODO_LOCAL" )
      Coil( "Signals".ProcessInterlock_APLC_Input[1].ModezoneInterlock_APLC_Input[2].StationInterlock_APLC_Input[16].PositionInterlock_APLC_Input[1].EquipmentInterlock_APLC_Input[1].SignalInterlock_APLC_Input[2] )
   END_RUNG
   RUNG wire#powerrail
      Contact( "Get_Cabine"."PORTAS CABINE" )
      I_Contact( "BYPASS_MOD_2" )
      I_Contact( "BYPASS_GERAL" )
      I_Contact( "BYPASS_CABINE_EM_MODO_LOCAL" )
      Coil( "Signals".ProcessInterlock_APLC_Input[1].ModezoneInterlock_APLC_Input[2].StationInterlock_APLC_Input[16].PositionInterlock_APLC_Input[1].EquipmentInterlock_APLC_Input[1].SignalInterlock_APLC_Input[3] )
   END_RUNG
   RUNG wire#powerrail
      Contact( "Get_Cabine".ROBO )
      I_Contact( "BYPASS_MOD_2" )
      I_Contact( "BYPASS_GERAL" )
      I_Contact( "BYPASS_CABINE_EM_MODO_LOCAL" )
      Coil( "Signals".ProcessInterlock_APLC_Input[1].ModezoneInterlock_APLC_Input[2].StationInterlock_APLC_Input[16].PositionInterlock_APLC_Input[1].EquipmentInterlock_APLC_Input[1].SignalInterlock_APLC_Input[4] )
   END_RUNG
   RUNG wire#powerrail
      Contact( "Get_Cabine"."TALHA FORA DE POSIÇÃO" )
      I_Contact( "BYPASS_MOD_2" )
      I_Contact( "BYPASS_GERAL" )
      I_Contact( "BYPASS_CABINE_EM_MODO_LOCAL" )
      Coil( "Signals".ProcessInterlock_APLC_Input[1].ModezoneInterlock_APLC_Input[2].StationInterlock_APLC_Input[16].PositionInterlock_APLC_Input[1].EquipmentInterlock_APLC_Input[1].SignalInterlock_APLC_Input[5] )
   END_RUNG
   RUNG wire#powerrail
      Contact( "Get_Cabine"."CABINE NOK" )
      I_Contact( "Get_Cabine".ROBO )
      Contact( "Get_Cabine"."CONFIRMAÇÃO DE RECEITA" )
      I_Contact( "Get_Cabine"."SIGNAL RESERVED"[1].BOOL_2 )
      I_Contact( "BYPASS_MOD_2" )
      I_Contact( "BYPASS_GERAL" )
      I_Contact( "BYPASS_CABINE_EM_MODO_LOCAL" )
      Coil( "Signals".ProcessInterlock_APLC_Input[1].ModezoneInterlock_APLC_Input[2].StationInterlock_APLC_Input[16].PositionInterlock_APLC_Input[1].EquipmentInterlock_APLC_Input[1].SignalInterlock_APLC_Input[6] )
   END_RUNG
   RUNG wire#powerrail
      I_Contact( "Get_Cabine"."CONFIRMAÇÃO DE RECEITA" )
      I_Contact( "BYPASS_MOD_2" )
      I_Contact( "BYPASS_GERAL" )
      I_Contact( "BYPASS_CABINE_EM_MODO_LOCAL" )
      Coil( "Signals".ProcessInterlock_APLC_Input[1].ModezoneInterlock_APLC_Input[2].StationInterlock_APLC_Input[16].PositionInterlock_APLC_Input[1].EquipmentInterlock_APLC_Input[1].SignalInterlock_APLC_Input[7] )
   END_RUNG
   RUNG wire#powerrail
      Contact( "Get_Cabine"."TAKT LOCAL" )
      I_Contact( "BYPASS_MOD_2" )
      I_Contact( "BYPASS_GERAL" )
      I_Contact( "BYPASS_CABINE_EM_MODO_LOCAL" )
      Coil( "Signals".ProcessInterlock_APLC_Input[1].ModezoneInterlock_APLC_Input[2].StationInterlock_APLC_Input[16].PositionInterlock_APLC_Input[1].EquipmentInterlock_APLC_Input[1].SignalInterlock_APLC_Input[8] )
   END_RUNG
   RUNG wire#powerrail
      Contact( "Get_Cabine"."SIGNAL RESERVED"[1]."BOOL" )
      I_Contact( "BYPASS_MOD_2" )
      I_Contact( "BYPASS_GERAL" )
      I_Contact( "BYPASS_CABINE_EM_MODO_LOCAL" )
      Coil( "Signals".ProcessInterlock_APLC_Input[1].ModezoneInterlock_APLC_Input[2].StationInterlock_APLC_Input[16].PositionInterlock_APLC_Input[1].EquipmentInterlock_APLC_Input[2].SignalInterlock_APLC_Input[1] )
   END_RUNG
   RUNG wire#powerrail
      Contact( "Get_Cabine"."SIGNAL RESERVED"[1].BOOL_1 )
      I_Contact( "BYPASS_MOD_2" )
      I_Contact( "BYPASS_GERAL" )
      I_Contact( "BYPASS_CABINE_EM_MODO_LOCAL" )
      Coil( "Signals".ProcessInterlock_APLC_Input[1].ModezoneInterlock_APLC_Input[2].StationInterlock_APLC_Input[16].PositionInterlock_APLC_Input[1].EquipmentInterlock_APLC_Input[2].SignalInterlock_APLC_Input[2] )
   END_RUNG
   RUNG wire#powerrail
      Contact( "Get_Cabine"."SIGNAL RESERVED"[1].BOOL_2 )
      I_Contact( "BYPASS_MOD_2" )
      I_Contact( "BYPASS_GERAL" )
      I_Contact( "BYPASS_CABINE_EM_MODO_LOCAL" )
      Coil( "Signals".ProcessInterlock_APLC_Input[1].ModezoneInterlock_APLC_Input[2].StationInterlock_APLC_Input[16].PositionInterlock_APLC_Input[1].EquipmentInterlock_APLC_Input[2].SignalInterlock_APLC_Input[3] )
   END_RUNG
   RUNG wire#powerrail
      Contact( "Get_Cabine"."SIGNAL RESERVED"[1].BOOL_3 )
      I_Contact( "BYPASS_MOD_2" )
      I_Contact( "BYPASS_GERAL" )
      I_Contact( "BYPASS_CABINE_EM_MODO_LOCAL" )
      Coil( "Signals".ProcessInterlock_APLC_Input[1].ModezoneInterlock_APLC_Input[2].StationInterlock_APLC_Input[16].PositionInterlock_APLC_Input[1].EquipmentInterlock_APLC_Input[2].SignalInterlock_APLC_Input[4] )
   END_RUNG
   RUNG wire#powerrail
      Contact( "Get_Cabine"."SIGNAL RESERVED"[2]."BOOL" )
      I_Contact( "BYPASS_MOD_2" )
      I_Contact( "BYPASS_GERAL" )
      I_Contact( "BYPASS_CABINE_EM_MODO_LOCAL" )
      Coil( "Put Sinais de Interlock Main line"."GIRO CABINE" )
   END_RUNG
   RUNG wire#powerrail
      Contact( "Get_Cabine"."SIGNAL RESERVED"[2].BOOL_1 )
      I_Contact( "BYPASS_MOD_2" )
      I_Contact( "BYPASS_GERAL" )
      I_Contact( "BYPASS_CABINE_EM_MODO_LOCAL" )
      Coil( "Signals".ProcessInterlock_APLC_Input[1].ModezoneInterlock_APLC_Input[2].StationInterlock_APLC_Input[16].PositionInterlock_APLC_Input[1].EquipmentInterlock_APLC_Input[2].SignalInterlock_APLC_Input[5] )
   END_RUNG
   RUNG wire#powerrail
      Contact( "Put_cabine"."Modezone done cab" )
      wire#w1
      I_Contact( "Get_Cabine"."SIGNAL RESERVED"[2]."BOOL" )
      { S7_Templates := "time_type := Time" } "IEC_Timer_0_DB_12".TON(pt := T#10S, et =>)
      Coil( "Signals".ProcessInterlock_APLC_Input[1].ModezoneInterlock_APLC_Input[2].StationInterlock_APLC_Input[16].PositionInterlock_APLC_Input[1].EquipmentInterlock_APLC_Input[2].SignalInterlock_APLC_Input[6] )
   END_RUNG
   RUNG wire#powerrail
      Contact( "Get_Cabine"."SIGNAL RESERVED"[5]."BOOL" )
   END_RUNG wire#w1
   // the same network as SCL:
   "Signals".ProcessInterlock_APLC_Input[1].ModezoneInterlock_APLC_Input[2].StationInterlock_APLC_Input[16].PositionInterlock_APLC_Input[1].EquipmentInterlock_APLC_Input[1].SignalInterlock_APLC_Input[1] := "Get_Cabine".ANDON AND NOT "BYPASS_MOD_2" AND NOT "BYPASS_GERAL" AND NOT "BYPASS_CABINE_EM_MODO_LOCAL";
   "Signals".ProcessInterlock_APLC_Input[1].ModezoneInterlock_APLC_Input[2].StationInterlock_APLC_Input[16].PositionInterlock_APLC_Input[1].EquipmentInterlock_APLC_Input[1].SignalInterlock_APLC_Input[2] := "Get_Cabine".EMERGÊNCIA AND NOT "BYPASS_MOD_2" AND NOT "BYPASS_GERAL" AND NOT "BYPASS_CABINE_EM_MODO_LOCAL";
   "Signals".ProcessInterlock_APLC_Input[1].ModezoneInterlock_APLC_Input[2].StationInterlock_APLC_Input[16].PositionInterlock_APLC_Input[1].EquipmentInterlock_APLC_Input[1].SignalInterlock_APLC_Input[3] := "Get_Cabine"."PORTAS CABINE" AND NOT "BYPASS_MOD_2" AND NOT "BYPASS_GERAL" AND NOT "BYPASS_CABINE_EM_MODO_LOCAL";
   "Signals".ProcessInterlock_APLC_Input[1].ModezoneInterlock_APLC_Input[2].StationInterlock_APLC_Input[16].PositionInterlock_APLC_Input[1].EquipmentInterlock_APLC_Input[1].SignalInterlock_APLC_Input[4] := "Get_Cabine".ROBO AND NOT "BYPASS_MOD_2" AND NOT "BYPASS_GERAL" AND NOT "BYPASS_CABINE_EM_MODO_LOCAL";
   "Signals".ProcessInterlock_APLC_Input[1].ModezoneInterlock_APLC_Input[2].StationInterlock_APLC_Input[16].PositionInterlock_APLC_Input[1].EquipmentInterlock_APLC_Input[1].SignalInterlock_APLC_Input[5] := "Get_Cabine"."TALHA FORA DE POSIÇÃO" AND NOT "BYPASS_MOD_2" AND NOT "BYPASS_GERAL" AND NOT "BYPASS_CABINE_EM_MODO_LOCAL";
   "Signals".ProcessInterlock_APLC_Input[1].ModezoneInterlock_APLC_Input[2].StationInterlock_APLC_Input[16].PositionInterlock_APLC_Input[1].EquipmentInterlock_APLC_Input[1].SignalInterlock_APLC_Input[6] := "Get_Cabine"."CABINE NOK" AND NOT "Get_Cabine".ROBO AND "Get_Cabine"."CONFIRMAÇÃO DE RECEITA" AND NOT "Get_Cabine"."SIGNAL RESERVED"[1].BOOL_2 AND NOT "BYPASS_MOD_2" AND NOT "BYPASS_GERAL" AND NOT "BYPASS_CABINE_EM_MODO_LOCAL";
   "Signals".ProcessInterlock_APLC_Input[1].ModezoneInterlock_APLC_Input[2].StationInterlock_APLC_Input[16].PositionInterlock_APLC_Input[1].EquipmentInterlock_APLC_Input[1].SignalInterlock_APLC_Input[7] := NOT "Get_Cabine"."CONFIRMAÇÃO DE RECEITA" AND NOT "BYPASS_MOD_2" AND NOT "BYPASS_GERAL" AND NOT "BYPASS_CABINE_EM_MODO_LOCAL";
   "Signals".ProcessInterlock_APLC_Input[1].ModezoneInterlock_APLC_Input[2].StationInterlock_APLC_Input[16].PositionInterlock_APLC_Input[1].EquipmentInterlock_APLC_Input[1].SignalInterlock_APLC_Input[8] := "Get_Cabine"."TAKT LOCAL" AND NOT "BYPASS_MOD_2" AND NOT "BYPASS_GERAL" AND NOT "BYPASS_CABINE_EM_MODO_LOCAL";
   "Signals".ProcessInterlock_APLC_Input[1].ModezoneInterlock_APLC_Input[2].StationInterlock_APLC_Input[16].PositionInterlock_APLC_Input[1].EquipmentInterlock_APLC_Input[2].SignalInterlock_APLC_Input[1] := "Get_Cabine"."SIGNAL RESERVED"[1]."BOOL" AND NOT "BYPASS_MOD_2" AND NOT "BYPASS_GERAL" AND NOT "BYPASS_CABINE_EM_MODO_LOCAL";
   "Signals".ProcessInterlock_APLC_Input[1].ModezoneInterlock_APLC_Input[2].StationInterlock_APLC_Input[16].PositionInterlock_APLC_Input[1].EquipmentInterlock_APLC_Input[2].SignalInterlock_APLC_Input[2] := "Get_Cabine"."SIGNAL RESERVED"[1].BOOL_1 AND NOT "BYPASS_MOD_2" AND NOT "BYPASS_GERAL" AND NOT "BYPASS_CABINE_EM_MODO_LOCAL";
   "Signals".ProcessInterlock_APLC_Input[1].ModezoneInterlock_APLC_Input[2].StationInterlock_APLC_Input[16].PositionInterlock_APLC_Input[1].EquipmentInterlock_APLC_Input[2].SignalInterlock_APLC_Input[3] := "Get_Cabine"."SIGNAL RESERVED"[1].BOOL_2 AND NOT "BYPASS_MOD_2" AND NOT "BYPASS_GERAL" AND NOT "BYPASS_CABINE_EM_MODO_LOCAL";
   "Signals".ProcessInterlock_APLC_Input[1].ModezoneInterlock_APLC_Input[2].StationInterlock_APLC_Input[16].PositionInterlock_APLC_Input[1].EquipmentInterlock_APLC_Input[2].SignalInterlock_APLC_Input[4] := "Get_Cabine"."SIGNAL RESERVED"[1].BOOL_3 AND NOT "BYPASS_MOD_2" AND NOT "BYPASS_GERAL" AND NOT "BYPASS_CABINE_EM_MODO_LOCAL";
   "Put Sinais de Interlock Main line"."GIRO CABINE" := "Get_Cabine"."SIGNAL RESERVED"[2]."BOOL" AND NOT "BYPASS_MOD_2" AND NOT "BYPASS_GERAL" AND NOT "BYPASS_CABINE_EM_MODO_LOCAL";
   "Signals".ProcessInterlock_APLC_Input[1].ModezoneInterlock_APLC_Input[2].StationInterlock_APLC_Input[16].PositionInterlock_APLC_Input[1].EquipmentInterlock_APLC_Input[2].SignalInterlock_APLC_Input[5] := "Get_Cabine"."SIGNAL RESERVED"[2].BOOL_1 AND NOT "BYPASS_MOD_2" AND NOT "BYPASS_GERAL" AND NOT "BYPASS_CABINE_EM_MODO_LOCAL";
   "IEC_Timer_0_DB_12".TON(IN := ("Put_cabine"."Modezone done cab" OR "Get_Cabine"."SIGNAL RESERVED"[5]."BOOL") AND NOT "Get_Cabine"."SIGNAL RESERVED"[2]."BOOL",
                           PT := T#10S);
   "Signals".ProcessInterlock_APLC_Input[1].ModezoneInterlock_APLC_Input[2].StationInterlock_APLC_Input[16].PositionInterlock_APLC_Input[1].EquipmentInterlock_APLC_Input[2].SignalInterlock_APLC_Input[6] := "IEC_Timer_0_DB_12".Q;
END_REGION

REGION Network 31: SINAIS ENVIADOS PARA CABINE
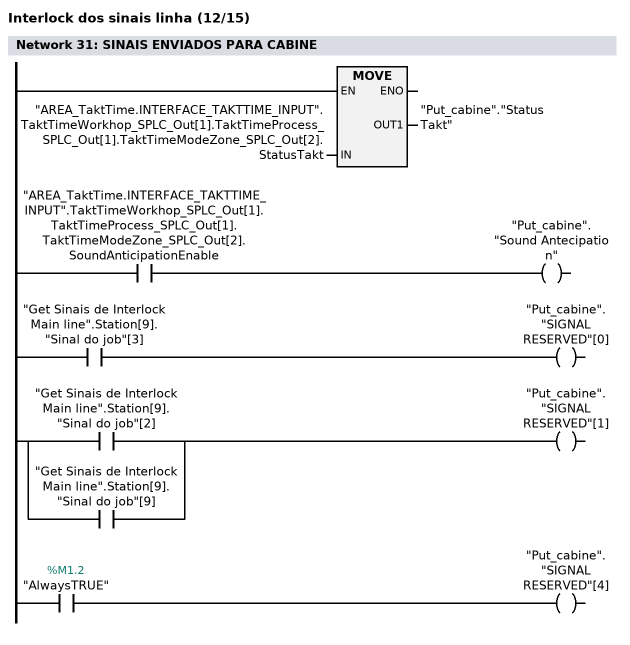
   RUNG wire#powerrail
      Move(in := "AREA_TaktTime.INTERFACE_TAKTTIME_INPUT".TaktTimeWorkhop_SPLC_Out[1].TaktTimeProcess_SPLC_Out[1].TaktTimeModeZone_SPLC_Out[2].StatusTakt, out1 => "Put_cabine"."Status Takt")
   END_RUNG
   RUNG wire#powerrail
      Contact( "AREA_TaktTime.INTERFACE_TAKTTIME_INPUT".TaktTimeWorkhop_SPLC_Out[1].TaktTimeProcess_SPLC_Out[1].TaktTimeModeZone_SPLC_Out[2].SoundAnticipationEnable )
      Coil( "Put_cabine"."Sound Antecipation" )
   END_RUNG
   RUNG wire#powerrail
      Contact( "Get Sinais de Interlock Main line".Station[9]."Sinal do job"[3] )
      Coil( "Put_cabine"."SIGNAL RESERVED"[0] )
   END_RUNG
   RUNG wire#powerrail
      Contact( "Get Sinais de Interlock Main line".Station[9]."Sinal do job"[2] )
      wire#w1
      Coil( "Put_cabine"."SIGNAL RESERVED"[1] )
   END_RUNG
   RUNG wire#powerrail
      Contact( "Get Sinais de Interlock Main line".Station[9]."Sinal do job"[9] )
   END_RUNG wire#w1
   RUNG wire#powerrail
      Contact( "AlwaysTRUE" )
      Coil( "Put_cabine"."SIGNAL RESERVED"[4] )
   END_RUNG
   // the same network as SCL:
   "Put_cabine"."Status Takt" := "AREA_TaktTime.INTERFACE_TAKTTIME_INPUT".TaktTimeWorkhop_SPLC_Out[1].TaktTimeProcess_SPLC_Out[1].TaktTimeModeZone_SPLC_Out[2].StatusTakt;
   "Put_cabine"."Sound Antecipation" := "AREA_TaktTime.INTERFACE_TAKTTIME_INPUT".TaktTimeWorkhop_SPLC_Out[1].TaktTimeProcess_SPLC_Out[1].TaktTimeModeZone_SPLC_Out[2].SoundAnticipationEnable;
   "Put_cabine"."SIGNAL RESERVED"[0] := "Get Sinais de Interlock Main line".Station[9]."Sinal do job"[3];
   "Put_cabine"."SIGNAL RESERVED"[1] := "Get Sinais de Interlock Main line".Station[9]."Sinal do job"[2] OR "Get Sinais de Interlock Main line".Station[9]."Sinal do job"[9];
   "Put_cabine"."SIGNAL RESERVED"[4] := "AlwaysTRUE";
END_REGION

REGION Network 32: Mod1 e 2 OK
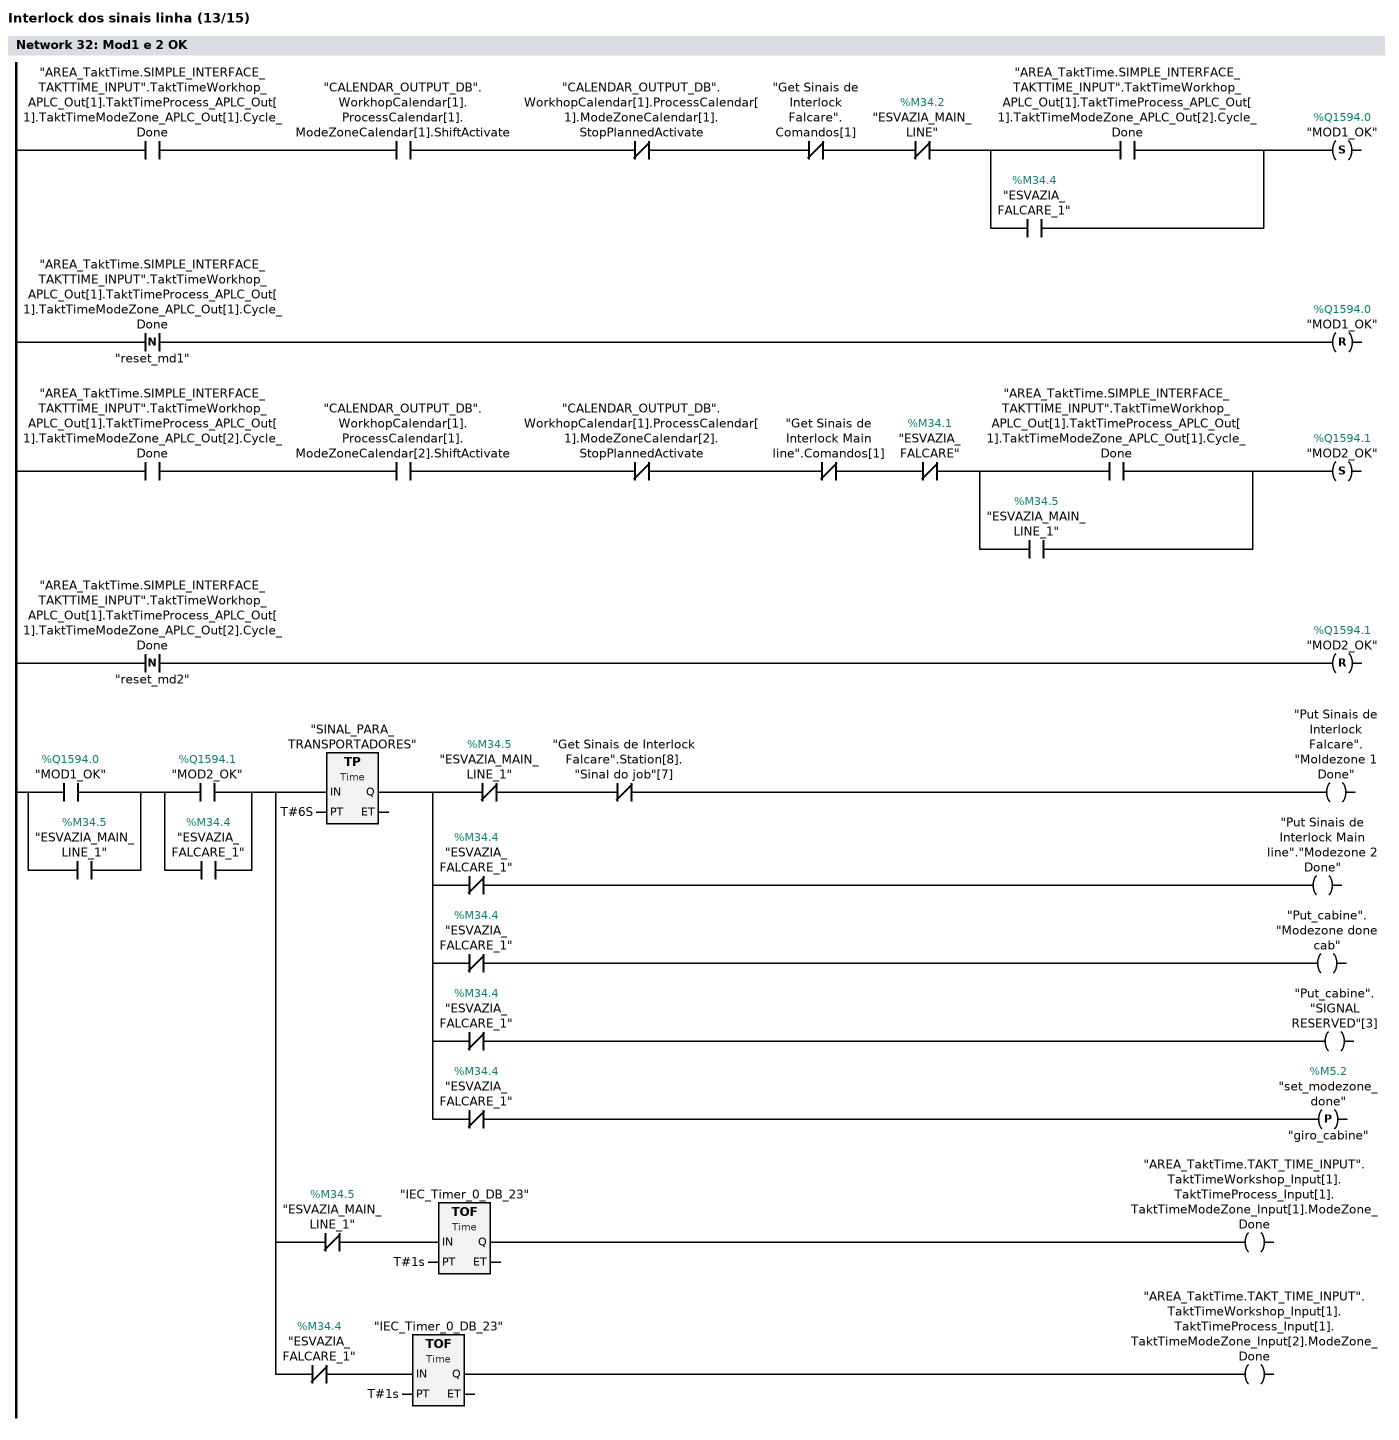
   IF "AREA_TaktTime.SIMPLE_INTERFACE_TAKTTIME_INPUT".TaktTimeWorkhop_APLC_Out[1].TaktTimeProcess_APLC_Out[1].TaktTimeModeZone_APLC_Out[1].Cycle_Done AND "CALENDAR_OUTPUT_DB".WorkhopCalendar[1].ProcessCalendar[1].ModeZoneCalendar[1].ShiftActivate AND NOT "CALENDAR_OUTPUT_DB".WorkhopCalendar[1].ProcessCalendar[1].ModeZoneCalendar[1].StopPlannedActivate AND NOT "Get Sinais de Interlock Falcare".Comandos[1] AND NOT "ESVAZIA_MAIN_LINE" AND ("AREA_TaktTime.SIMPLE_INTERFACE_TAKTTIME_INPUT".TaktTimeWorkhop_APLC_Out[1].TaktTimeProcess_APLC_Out[1].TaktTimeModeZone_APLC_Out[2].Cycle_Done OR "ESVAZIA_FALCARE_1") THEN
       "MOD1_OK" := TRUE;
   END_IF;
   #_w1 := NOT "AREA_TaktTime.SIMPLE_INTERFACE_TAKTTIME_INPUT".TaktTimeWorkhop_APLC_Out[1].TaktTimeProcess_APLC_Out[1].TaktTimeModeZone_APLC_Out[1].Cycle_Done AND "reset_md1";   // falling edge of "AREA_TaktTime.SIMPLE_INTERFACE_TAKTTIME_INPUT".TaktTimeWorkhop_APLC_Out[1].TaktTimeProcess_APLC_Out[1].TaktTimeModeZone_APLC_Out[1].Cycle_Done
   "reset_md1" := "AREA_TaktTime.SIMPLE_INTERFACE_TAKTTIME_INPUT".TaktTimeWorkhop_APLC_Out[1].TaktTimeProcess_APLC_Out[1].TaktTimeModeZone_APLC_Out[1].Cycle_Done;
   IF #_w1 THEN "MOD1_OK" := FALSE; END_IF;
   IF "AREA_TaktTime.SIMPLE_INTERFACE_TAKTTIME_INPUT".TaktTimeWorkhop_APLC_Out[1].TaktTimeProcess_APLC_Out[1].TaktTimeModeZone_APLC_Out[2].Cycle_Done AND "CALENDAR_OUTPUT_DB".WorkhopCalendar[1].ProcessCalendar[1].ModeZoneCalendar[2].ShiftActivate AND NOT "CALENDAR_OUTPUT_DB".WorkhopCalendar[1].ProcessCalendar[1].ModeZoneCalendar[2].StopPlannedActivate AND NOT "Get Sinais de Interlock Main line".Comandos[1] AND NOT "ESVAZIA_FALCARE" AND ("AREA_TaktTime.SIMPLE_INTERFACE_TAKTTIME_INPUT".TaktTimeWorkhop_APLC_Out[1].TaktTimeProcess_APLC_Out[1].TaktTimeModeZone_APLC_Out[1].Cycle_Done OR "ESVAZIA_MAIN_LINE_1") THEN
       "MOD2_OK" := TRUE;
   END_IF;
   #_w2 := NOT "AREA_TaktTime.SIMPLE_INTERFACE_TAKTTIME_INPUT".TaktTimeWorkhop_APLC_Out[1].TaktTimeProcess_APLC_Out[1].TaktTimeModeZone_APLC_Out[2].Cycle_Done AND "reset_md2";   // falling edge of "AREA_TaktTime.SIMPLE_INTERFACE_TAKTTIME_INPUT".TaktTimeWorkhop_APLC_Out[1].TaktTimeProcess_APLC_Out[1].TaktTimeModeZone_APLC_Out[2].Cycle_Done
   "reset_md2" := "AREA_TaktTime.SIMPLE_INTERFACE_TAKTTIME_INPUT".TaktTimeWorkhop_APLC_Out[1].TaktTimeProcess_APLC_Out[1].TaktTimeModeZone_APLC_Out[2].Cycle_Done;
   IF #_w2 THEN "MOD2_OK" := FALSE; END_IF;
   #_w3 := ("MOD1_OK" OR "ESVAZIA_MAIN_LINE_1") AND ("MOD2_OK" OR "ESVAZIA_FALCARE_1");
   "SINAL_PARA_TRANSPORTADORES".TP(IN := #_w3, PT := T#6S);
   "Put Sinais de Interlock Falcare"."Moldezone 1 Done" := "SINAL_PARA_TRANSPORTADORES".Q AND NOT "ESVAZIA_MAIN_LINE_1" AND NOT "Get Sinais de Interlock Falcare".Station[8]."Sinal do job"[7];
   "Put Sinais de Interlock Main line"."Modezone 2 Done" := "SINAL_PARA_TRANSPORTADORES".Q AND NOT "ESVAZIA_FALCARE_1";
   "Put_cabine"."Modezone done cab" := "SINAL_PARA_TRANSPORTADORES".Q AND NOT "ESVAZIA_FALCARE_1";
   "Put_cabine"."SIGNAL RESERVED"[3] := "SINAL_PARA_TRANSPORTADORES".Q AND NOT "ESVAZIA_FALCARE_1";
   #_w4 := "SINAL_PARA_TRANSPORTADORES".Q AND NOT "ESVAZIA_FALCARE_1";
   "set_modezone_done" := #_w4 AND NOT "giro_cabine";   // rising edge
   "giro_cabine" := #_w4;
   "IEC_Timer_0_DB_23".TOF(IN := #_w3 AND NOT "ESVAZIA_MAIN_LINE_1", PT := T#1s);
   "AREA_TaktTime.TAKT_TIME_INPUT".TaktTimeWorkshop_Input[1].TaktTimeProcess_Input[1].TaktTimeModeZone_Input[1].ModeZone_Done := "IEC_Timer_0_DB_23".Q;
   "IEC_Timer_0_DB_23".TOF(IN := #_w3 AND NOT "ESVAZIA_FALCARE_1", PT := T#1s);
   "AREA_TaktTime.TAKT_TIME_INPUT".TaktTimeWorkshop_Input[1].TaktTimeProcess_Input[1].TaktTimeModeZone_Input[2].ModeZone_Done := "IEC_Timer_0_DB_23".Q;
END_REGION

REGION Network 33: LIBERAÇÃO DE TURNO ATIVO PARA TRANSPORTADORES FALCARE E MAIN LINE / CABINE DE PINTURA
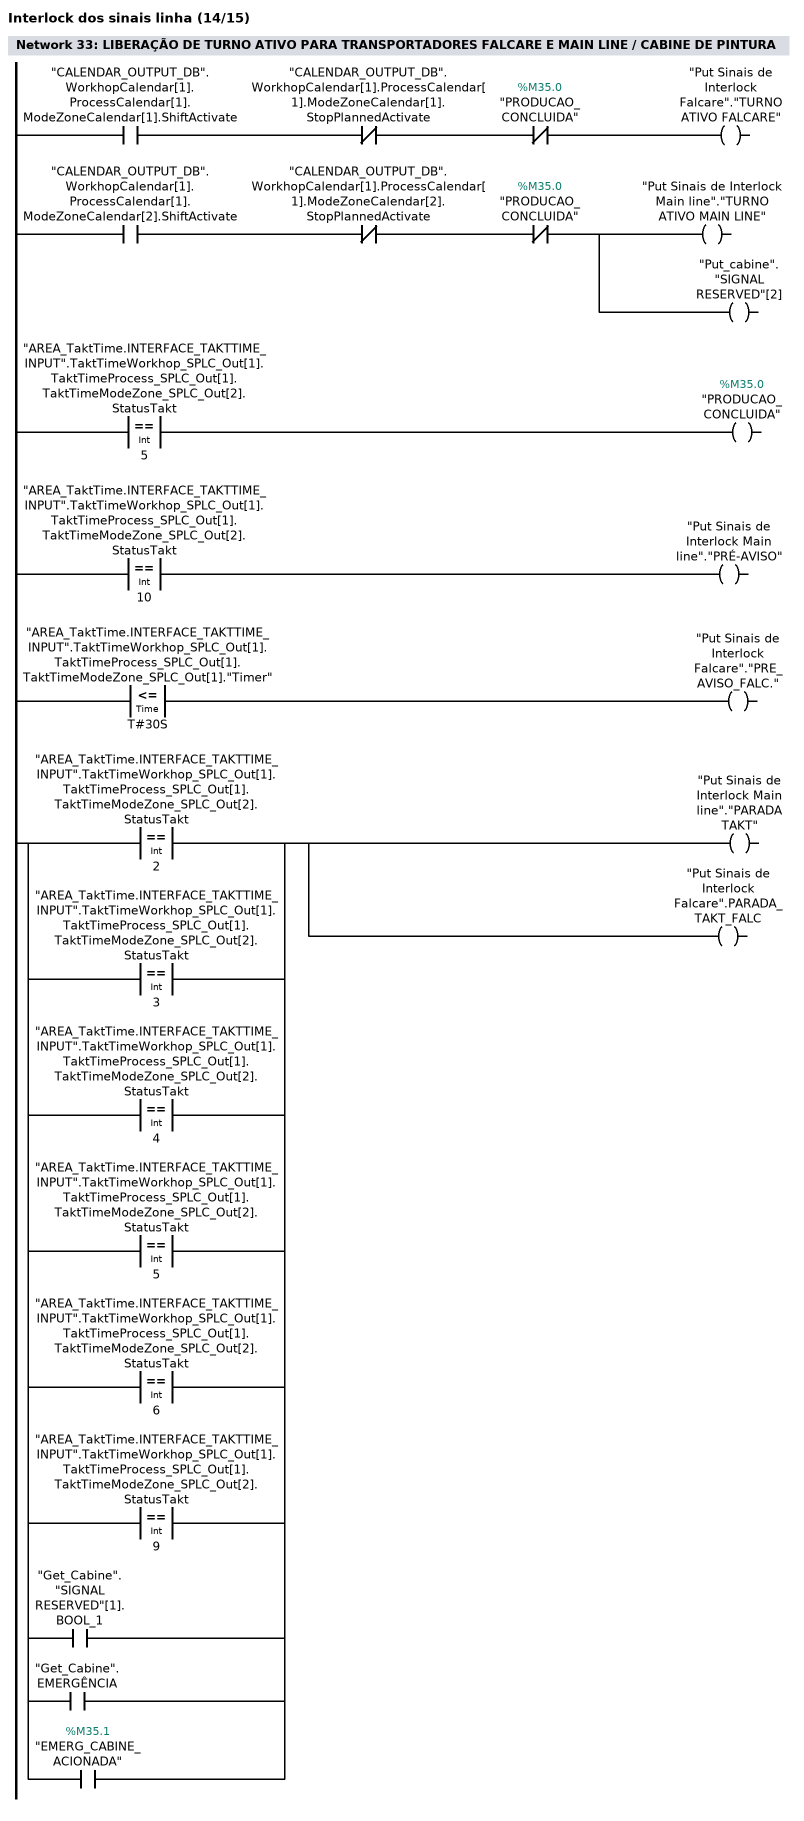
   RUNG wire#powerrail
      Contact( "CALENDAR_OUTPUT_DB".WorkhopCalendar[1].ProcessCalendar[1].ModeZoneCalendar[1].ShiftActivate )
      I_Contact( "CALENDAR_OUTPUT_DB".WorkhopCalendar[1].ProcessCalendar[1].ModeZoneCalendar[1].StopPlannedActivate )
      I_Contact( "PRODUCAO_CONCLUIDA" )
      Coil( "Put Sinais de Interlock Falcare"."TURNO ATIVO FALCARE" )
   END_RUNG
   RUNG wire#powerrail
      Contact( "CALENDAR_OUTPUT_DB".WorkhopCalendar[1].ProcessCalendar[1].ModeZoneCalendar[2].ShiftActivate )
      I_Contact( "CALENDAR_OUTPUT_DB".WorkhopCalendar[1].ProcessCalendar[1].ModeZoneCalendar[2].StopPlannedActivate )
      I_Contact( "PRODUCAO_CONCLUIDA" )
      wire#w1
      Coil( "Put Sinais de Interlock Main line"."TURNO ATIVO MAIN LINE" )
   END_RUNG
   RUNG wire#w1
      Coil( "Put_cabine"."SIGNAL RESERVED"[2] )
   END_RUNG
   RUNG wire#powerrail
      { S7_Templates := "SrcType := Int" } EQ_Contact(in1 := "AREA_TaktTime.INTERFACE_TAKTTIME_INPUT".TaktTimeWorkhop_SPLC_Out[1].TaktTimeProcess_SPLC_Out[1].TaktTimeModeZone_SPLC_Out[2].StatusTakt, in2 := 5)
      Coil( "PRODUCAO_CONCLUIDA" )
   END_RUNG
   RUNG wire#powerrail
      { S7_Templates := "SrcType := Int" } EQ_Contact(in1 := "AREA_TaktTime.INTERFACE_TAKTTIME_INPUT".TaktTimeWorkhop_SPLC_Out[1].TaktTimeProcess_SPLC_Out[1].TaktTimeModeZone_SPLC_Out[2].StatusTakt, in2 := 10)
      Coil( "Put Sinais de Interlock Main line"."PRÉ-AVISO" )
   END_RUNG
   RUNG wire#powerrail
      { S7_Templates := "SrcType := Time" } LE_Contact(in1 := "AREA_TaktTime.INTERFACE_TAKTTIME_INPUT".TaktTimeWorkhop_SPLC_Out[1].TaktTimeProcess_SPLC_Out[1].TaktTimeModeZone_SPLC_Out[1]."Timer", in2 := T#30S)
      Coil( "Put Sinais de Interlock Falcare"."PRE_AVISO_FALC." )
   END_RUNG
   RUNG wire#powerrail
      { S7_Templates := "SrcType := Int" } EQ_Contact(in1 := "AREA_TaktTime.INTERFACE_TAKTTIME_INPUT".TaktTimeWorkhop_SPLC_Out[1].TaktTimeProcess_SPLC_Out[1].TaktTimeModeZone_SPLC_Out[2].StatusTakt, in2 := 2)
      wire#w2
      Coil( "Put Sinais de Interlock Main line"."PARADA TAKT" )
   END_RUNG
   RUNG wire#powerrail
      { S7_Templates := "SrcType := Int" } EQ_Contact(in1 := "AREA_TaktTime.INTERFACE_TAKTTIME_INPUT".TaktTimeWorkhop_SPLC_Out[1].TaktTimeProcess_SPLC_Out[1].TaktTimeModeZone_SPLC_Out[2].StatusTakt, in2 := 3)
   END_RUNG wire#w2
   RUNG wire#powerrail
      { S7_Templates := "SrcType := Int" } EQ_Contact(in1 := "AREA_TaktTime.INTERFACE_TAKTTIME_INPUT".TaktTimeWorkhop_SPLC_Out[1].TaktTimeProcess_SPLC_Out[1].TaktTimeModeZone_SPLC_Out[2].StatusTakt, in2 := 4)
   END_RUNG wire#w2
   RUNG wire#powerrail
      { S7_Templates := "SrcType := Int" } EQ_Contact(in1 := "AREA_TaktTime.INTERFACE_TAKTTIME_INPUT".TaktTimeWorkhop_SPLC_Out[1].TaktTimeProcess_SPLC_Out[1].TaktTimeModeZone_SPLC_Out[2].StatusTakt, in2 := 5)
   END_RUNG wire#w2
   RUNG wire#powerrail
      { S7_Templates := "SrcType := Int" } EQ_Contact(in1 := "AREA_TaktTime.INTERFACE_TAKTTIME_INPUT".TaktTimeWorkhop_SPLC_Out[1].TaktTimeProcess_SPLC_Out[1].TaktTimeModeZone_SPLC_Out[2].StatusTakt, in2 := 6)
   END_RUNG wire#w2
   RUNG wire#powerrail
      { S7_Templates := "SrcType := Int" } EQ_Contact(in1 := "AREA_TaktTime.INTERFACE_TAKTTIME_INPUT".TaktTimeWorkhop_SPLC_Out[1].TaktTimeProcess_SPLC_Out[1].TaktTimeModeZone_SPLC_Out[2].StatusTakt, in2 := 9)
   END_RUNG wire#w2
   RUNG wire#powerrail
      Contact( "Get_Cabine"."SIGNAL RESERVED"[1].BOOL_1 )
   END_RUNG wire#w2
   RUNG wire#powerrail
      Contact( "Get_Cabine".EMERGÊNCIA )
   END_RUNG wire#w2
   RUNG wire#powerrail
      Contact( "EMERG_CABINE_ACIONADA" )
   END_RUNG wire#w2
   RUNG wire#w2
      Coil( "Put Sinais de Interlock Falcare".PARADA_TAKT_FALC )
   END_RUNG
   // the same network as SCL:
   "Put Sinais de Interlock Falcare"."TURNO ATIVO FALCARE" := "CALENDAR_OUTPUT_DB".WorkhopCalendar[1].ProcessCalendar[1].ModeZoneCalendar[1].ShiftActivate AND NOT "CALENDAR_OUTPUT_DB".WorkhopCalendar[1].ProcessCalendar[1].ModeZoneCalendar[1].StopPlannedActivate AND NOT "PRODUCAO_CONCLUIDA";
   "Put Sinais de Interlock Main line"."TURNO ATIVO MAIN LINE" := "CALENDAR_OUTPUT_DB".WorkhopCalendar[1].ProcessCalendar[1].ModeZoneCalendar[2].ShiftActivate AND NOT "CALENDAR_OUTPUT_DB".WorkhopCalendar[1].ProcessCalendar[1].ModeZoneCalendar[2].StopPlannedActivate AND NOT "PRODUCAO_CONCLUIDA";
   "Put_cabine"."SIGNAL RESERVED"[2] := "Put Sinais de Interlock Main line"."TURNO ATIVO MAIN LINE";
   "PRODUCAO_CONCLUIDA" := "AREA_TaktTime.INTERFACE_TAKTTIME_INPUT".TaktTimeWorkhop_SPLC_Out[1].TaktTimeProcess_SPLC_Out[1].TaktTimeModeZone_SPLC_Out[2].StatusTakt = 5;
   "Put Sinais de Interlock Main line"."PRÉ-AVISO" := "AREA_TaktTime.INTERFACE_TAKTTIME_INPUT".TaktTimeWorkhop_SPLC_Out[1].TaktTimeProcess_SPLC_Out[1].TaktTimeModeZone_SPLC_Out[2].StatusTakt = 10;
   "Put Sinais de Interlock Falcare"."PRE_AVISO_FALC." := "AREA_TaktTime.INTERFACE_TAKTTIME_INPUT".TaktTimeWorkhop_SPLC_Out[1].TaktTimeProcess_SPLC_Out[1].TaktTimeModeZone_SPLC_Out[1]."Timer" <= T#30S;
   "Put Sinais de Interlock Main line"."PARADA TAKT" := ("AREA_TaktTime.INTERFACE_TAKTTIME_INPUT".TaktTimeWorkhop_SPLC_Out[1].TaktTimeProcess_SPLC_Out[1].TaktTimeModeZone_SPLC_Out[2].StatusTakt = 2) OR ("AREA_TaktTime.INTERFACE_TAKTTIME_INPUT".TaktTimeWorkhop_SPLC_Out[1].TaktTimeProcess_SPLC_Out[1].TaktTimeModeZone_SPLC_Out[2].StatusTakt = 3) OR ("AREA_TaktTime.INTERFACE_TAKTTIME_INPUT".TaktTimeWorkhop_SPLC_Out[1].TaktTimeProcess_SPLC_Out[1].TaktTimeModeZone_SPLC_Out[2].StatusTakt = 4) OR ("AREA_TaktTime.INTERFACE_TAKTTIME_INPUT".TaktTimeWorkhop_SPLC_Out[1].TaktTimeProcess_SPLC_Out[1].TaktTimeModeZone_SPLC_Out[2].StatusTakt = 5) OR ("AREA_TaktTime.INTERFACE_TAKTTIME_INPUT".TaktTimeWorkhop_SPLC_Out[1].TaktTimeProcess_SPLC_Out[1].TaktTimeModeZone_SPLC_Out[2].StatusTakt = 6) OR ("AREA_TaktTime.INTERFACE_TAKTTIME_INPUT".TaktTimeWorkhop_SPLC_Out[1].TaktTimeProcess_SPLC_Out[1].TaktTimeModeZone_SPLC_Out[2].StatusTakt = 9) OR "Get_Cabine"."SIGNAL RESERVED"[1].BOOL_1 OR "Get_Cabine".EMERGÊNCIA OR "EMERG_CABINE_ACIONADA";
   "Put Sinais de Interlock Falcare".PARADA_TAKT_FALC := "Put Sinais de Interlock Main line"."PARADA TAKT";
END_REGION

REGION Network 34: LIFE BIT PARA TRANSPORTADORES
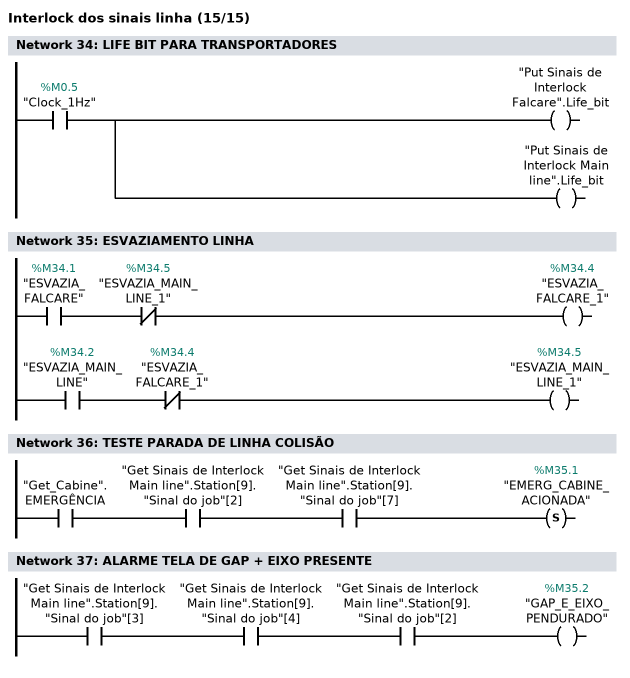
   RUNG wire#powerrail
      Contact( "Clock_1Hz" )
      wire#w1
      Coil( "Put Sinais de Interlock Falcare".Life_bit )
   END_RUNG
   RUNG wire#w1
      Coil( "Put Sinais de Interlock Main line".Life_bit )
   END_RUNG
   // the same network as SCL:
   "Put Sinais de Interlock Falcare".Life_bit := "Clock_1Hz";
   "Put Sinais de Interlock Main line".Life_bit := "Clock_1Hz";
END_REGION

REGION Network 35: ESVAZIAMENTO LINHA
   RUNG wire#powerrail
      Contact( "ESVAZIA_FALCARE" )
      I_Contact( "ESVAZIA_MAIN_LINE_1" )
      Coil( "ESVAZIA_FALCARE_1" )
   END_RUNG
   RUNG wire#powerrail
      Contact( "ESVAZIA_MAIN_LINE" )
      I_Contact( "ESVAZIA_FALCARE_1" )
      Coil( "ESVAZIA_MAIN_LINE_1" )
   END_RUNG
   // the same network as SCL:
   "ESVAZIA_FALCARE_1" := "ESVAZIA_FALCARE" AND NOT "ESVAZIA_MAIN_LINE_1";
   "ESVAZIA_MAIN_LINE_1" := "ESVAZIA_MAIN_LINE" AND NOT "ESVAZIA_FALCARE_1";
END_REGION

REGION Network 36: TESTE PARADA DE LINHA COLISÃO
   RUNG wire#powerrail
      Contact( "Get_Cabine".EMERGÊNCIA )
      Contact( "Get Sinais de Interlock Main line".Station[9]."Sinal do job"[2] )
      Contact( "Get Sinais de Interlock Main line".Station[9]."Sinal do job"[7] )
      S_Coil( "EMERG_CABINE_ACIONADA" )
   END_RUNG
   // the same network as SCL:
   IF "Get_Cabine".EMERGÊNCIA AND "Get Sinais de Interlock Main line".Station[9]."Sinal do job"[2] AND "Get Sinais de Interlock Main line".Station[9]."Sinal do job"[7] THEN
       "EMERG_CABINE_ACIONADA" := TRUE;
   END_IF;
END_REGION

REGION Network 37: ALARME TELA DE GAP + EIXO PRESENTE
   RUNG wire#powerrail
      Contact( "Get Sinais de Interlock Main line".Station[9]."Sinal do job"[3] )
      Contact( "Get Sinais de Interlock Main line".Station[9]."Sinal do job"[4] )
      Contact( "Get Sinais de Interlock Main line".Station[9]."Sinal do job"[2] )
      Coil( "GAP_E_EIXO_PENDURADO" )
   END_RUNG
   // the same network as SCL:
   "GAP_E_EIXO_PENDURADO" := "Get Sinais de Interlock Main line".Station[9]."Sinal do job"[3] AND "Get Sinais de Interlock Main line".Station[9]."Sinal do job"[4] AND "Get Sinais de Interlock Main line".Station[9]."Sinal do job"[2];
END_REGION

REGION Network 38 (SCL): SEM JOB POKA YOKE P100 ORING MAP
   IF "EQUIPAMENTOS_RECIPE_POS_TAKT".EQUIPAMENTOS[17].RECIPE = 'ETRCALIP01' THEN
   "Put Sinais de Interlock Main line".RESERVED_4 := TRUE;
   ELSIF "BORDA_MD2".Q THEN
       "Put Sinais de Interlock Main line".RESERVED_4 := FALSE;
   END_IF;
END_REGION
END_FUNCTION

FUNCTION "RESET_MODZONES" : Void   // FC10, LAD
{ S7_Optimized_Access := 'TRUE' }
// stored: SetENOAutomatically false
BEGIN

REGION Network 1: RESET MOD 1
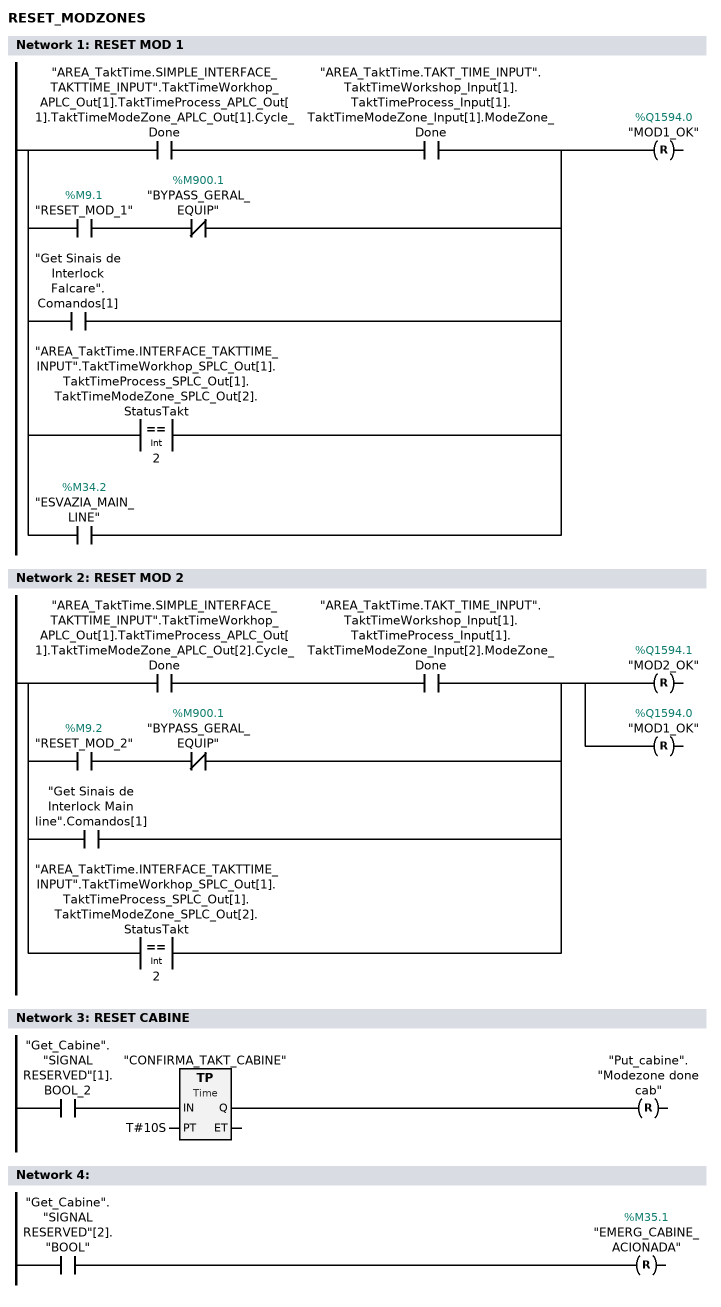
   RUNG wire#powerrail
      Contact( "AREA_TaktTime.SIMPLE_INTERFACE_TAKTTIME_INPUT".TaktTimeWorkhop_APLC_Out[1].TaktTimeProcess_APLC_Out[1].TaktTimeModeZone_APLC_Out[1].Cycle_Done )
      Contact( "AREA_TaktTime.TAKT_TIME_INPUT".TaktTimeWorkshop_Input[1].TaktTimeProcess_Input[1].TaktTimeModeZone_Input[1].ModeZone_Done )
      wire#w1
      R_Coil( "MOD1_OK" )
   END_RUNG
   RUNG wire#powerrail
      Contact( "RESET_MOD_1" )
      I_Contact( "BYPASS_GERAL_EQUIP" )
   END_RUNG wire#w1
   RUNG wire#powerrail
      Contact( "Get Sinais de Interlock Falcare".Comandos[1] )
   END_RUNG wire#w1
   RUNG wire#powerrail
      { S7_Templates := "SrcType := Int" } EQ_Contact(in1 := "AREA_TaktTime.INTERFACE_TAKTTIME_INPUT".TaktTimeWorkhop_SPLC_Out[1].TaktTimeProcess_SPLC_Out[1].TaktTimeModeZone_SPLC_Out[2].StatusTakt, in2 := 2)
   END_RUNG wire#w1
   RUNG wire#powerrail
      Contact( "ESVAZIA_MAIN_LINE" )
   END_RUNG wire#w1
   // the same network as SCL:
   IF ("AREA_TaktTime.SIMPLE_INTERFACE_TAKTTIME_INPUT".TaktTimeWorkhop_APLC_Out[1].TaktTimeProcess_APLC_Out[1].TaktTimeModeZone_APLC_Out[1].Cycle_Done AND "AREA_TaktTime.TAKT_TIME_INPUT".TaktTimeWorkshop_Input[1].TaktTimeProcess_Input[1].TaktTimeModeZone_Input[1].ModeZone_Done) OR ("RESET_MOD_1" AND NOT "BYPASS_GERAL_EQUIP") OR "Get Sinais de Interlock Falcare".Comandos[1] OR ("AREA_TaktTime.INTERFACE_TAKTTIME_INPUT".TaktTimeWorkhop_SPLC_Out[1].TaktTimeProcess_SPLC_Out[1].TaktTimeModeZone_SPLC_Out[2].StatusTakt = 2) OR "ESVAZIA_MAIN_LINE" THEN
       "MOD1_OK" := FALSE;
   END_IF;
END_REGION

REGION Network 2: RESET MOD 2
   RUNG wire#powerrail
      Contact( "AREA_TaktTime.SIMPLE_INTERFACE_TAKTTIME_INPUT".TaktTimeWorkhop_APLC_Out[1].TaktTimeProcess_APLC_Out[1].TaktTimeModeZone_APLC_Out[2].Cycle_Done )
      Contact( "AREA_TaktTime.TAKT_TIME_INPUT".TaktTimeWorkshop_Input[1].TaktTimeProcess_Input[1].TaktTimeModeZone_Input[2].ModeZone_Done )
      wire#w1
      R_Coil( "MOD2_OK" )
   END_RUNG
   RUNG wire#powerrail
      Contact( "RESET_MOD_2" )
      I_Contact( "BYPASS_GERAL_EQUIP" )
   END_RUNG wire#w1
   RUNG wire#powerrail
      Contact( "Get Sinais de Interlock Main line".Comandos[1] )
   END_RUNG wire#w1
   RUNG wire#powerrail
      { S7_Templates := "SrcType := Int" } EQ_Contact(in1 := "AREA_TaktTime.INTERFACE_TAKTTIME_INPUT".TaktTimeWorkhop_SPLC_Out[1].TaktTimeProcess_SPLC_Out[1].TaktTimeModeZone_SPLC_Out[2].StatusTakt, in2 := 2)
   END_RUNG wire#w1
   RUNG wire#w1
      R_Coil( "MOD1_OK" )
   END_RUNG
   // the same network as SCL:
   IF ("AREA_TaktTime.SIMPLE_INTERFACE_TAKTTIME_INPUT".TaktTimeWorkhop_APLC_Out[1].TaktTimeProcess_APLC_Out[1].TaktTimeModeZone_APLC_Out[2].Cycle_Done AND "AREA_TaktTime.TAKT_TIME_INPUT".TaktTimeWorkshop_Input[1].TaktTimeProcess_Input[1].TaktTimeModeZone_Input[2].ModeZone_Done) OR ("RESET_MOD_2" AND NOT "BYPASS_GERAL_EQUIP") OR "Get Sinais de Interlock Main line".Comandos[1] OR ("AREA_TaktTime.INTERFACE_TAKTTIME_INPUT".TaktTimeWorkhop_SPLC_Out[1].TaktTimeProcess_SPLC_Out[1].TaktTimeModeZone_SPLC_Out[2].StatusTakt = 2) THEN
       "MOD2_OK" := FALSE;
       "MOD1_OK" := FALSE;
   END_IF;
END_REGION

REGION Network 3: RESET CABINE
   RUNG wire#powerrail
      Contact( "Get_Cabine"."SIGNAL RESERVED"[1].BOOL_2 )
      { S7_Templates := "time_type := Time" } "CONFIRMA_TAKT_CABINE".TP(pt := T#10S, et =>)
      R_Coil( "Put_cabine"."Modezone done cab" )
   END_RUNG
   // the same network as SCL:
   "CONFIRMA_TAKT_CABINE".TP(IN := "Get_Cabine"."SIGNAL RESERVED"[1].BOOL_2, PT := T#10S);
   IF "CONFIRMA_TAKT_CABINE".Q THEN "Put_cabine"."Modezone done cab" := FALSE; END_IF;
END_REGION

REGION Network 4
   RUNG wire#powerrail
      Contact( "Get_Cabine"."SIGNAL RESERVED"[2]."BOOL" )
      R_Coil( "EMERG_CABINE_ACIONADA" )
   END_RUNG
   // the same network as SCL:
   IF "Get_Cabine"."SIGNAL RESERVED"[2]."BOOL" THEN "EMERG_CABINE_ACIONADA" := FALSE; END_IF;
END_REGION
END_FUNCTION

FUNCTION "VALIDACAO_ DOS_MODEZONES_ETR" : Void   // FC11, LAD
{ S7_Optimized_Access := 'TRUE' }
// stored: SetENOAutomatically false
   VAR_TEMP
      TESTE_1 : Bool;
      INDEX_STATION : Int;
      INDEX_POSITION : Int;
      INDEX_EQUIPMENT : Int;
      INDEX_SIGNAL : Int;
      leandro : Bool;
      index_positon_md1 : Int;
      index_equipament_md1 : Int;
      index_sinal_md1 : Int;
      POP_ID : String;
      BORDA : Bool;
      INDEX_CLEAN : Int;
      INDEX_FILA : Int;
      BORDA_1 : Bool;
      INDEX_SIGNAL1 : Int;
      INDEX_SIGNAL2 : Int;
      INDEX_VERIFICA : Int;
      barreira_invadida : Bool;
      aciona_buzzer : Bool;
      aciona_lampada_vermelha : Bool;
      aciona_lampada_verde : Bool;
      INTERLOCKS_MD1 : Bool;
      STATION : Int;
      SIGNAL : Int;
      EQUIPMENT : Int;
      count_LD : Bool;
      count_LE : Bool;
   END_VAR
   VAR_TEMP   // added for the SCL form of the ladder/FBD networks
      _w1 : Bool;
      _w2 : Bool;
   END_VAR
BEGIN

REGION Network 1: Buzzer
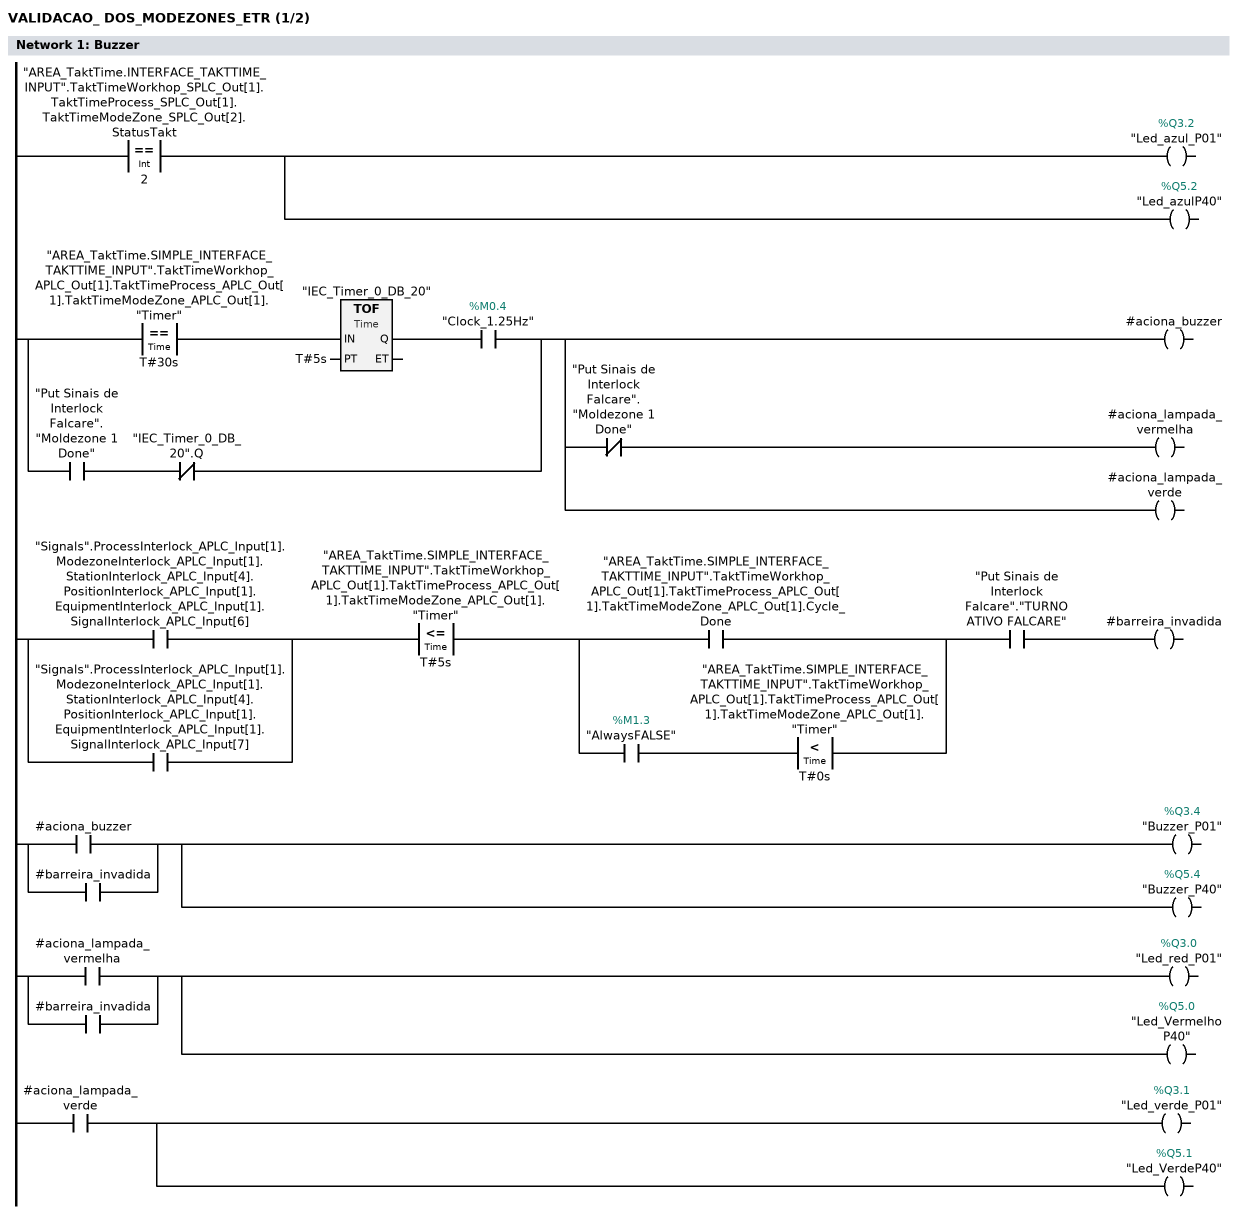
   RUNG wire#powerrail
      { S7_Templates := "SrcType := Int" } EQ_Contact(in1 := "AREA_TaktTime.INTERFACE_TAKTTIME_INPUT".TaktTimeWorkhop_SPLC_Out[1].TaktTimeProcess_SPLC_Out[1].TaktTimeModeZone_SPLC_Out[2].StatusTakt, in2 := 2)
      wire#w1
      Coil( "Led_azul_P01" )
   END_RUNG
   RUNG wire#w1
      Coil( "Led_azulP40" )
   END_RUNG
   RUNG wire#powerrail
      { S7_Templates := "SrcType := Time" } EQ_Contact(in1 := "AREA_TaktTime.SIMPLE_INTERFACE_TAKTTIME_INPUT".TaktTimeWorkhop_APLC_Out[1].TaktTimeProcess_APLC_Out[1].TaktTimeModeZone_APLC_Out[1]."Timer", in2 := T#30s)
      { S7_Templates := "time_type := Time" } "IEC_Timer_0_DB_20".TOF(pt := T#5s, et =>)
      Contact( "Clock_1.25Hz" )
      wire#w2
      Coil( #aciona_buzzer )
   END_RUNG
   RUNG wire#powerrail
      Contact( "Put Sinais de Interlock Falcare"."Moldezone 1 Done" )
      I_Contact( "IEC_Timer_0_DB_20".Q )
   END_RUNG wire#w2
   RUNG wire#w2
      I_Contact( "Put Sinais de Interlock Falcare"."Moldezone 1 Done" )
      Coil( #aciona_lampada_vermelha )
   END_RUNG
   RUNG wire#w2
      Coil( #aciona_lampada_verde )
   END_RUNG
   RUNG wire#powerrail
      Contact( "Signals".ProcessInterlock_APLC_Input[1].ModezoneInterlock_APLC_Input[1].StationInterlock_APLC_Input[4].PositionInterlock_APLC_Input[1].EquipmentInterlock_APLC_Input[1].SignalInterlock_APLC_Input[6] )
      wire#w3
      { S7_Templates := "SrcType := Time" } LE_Contact(in1 := "AREA_TaktTime.SIMPLE_INTERFACE_TAKTTIME_INPUT".TaktTimeWorkhop_APLC_Out[1].TaktTimeProcess_APLC_Out[1].TaktTimeModeZone_APLC_Out[1]."Timer", in2 := T#5s)
      wire#w4
      Contact( "AREA_TaktTime.SIMPLE_INTERFACE_TAKTTIME_INPUT".TaktTimeWorkhop_APLC_Out[1].TaktTimeProcess_APLC_Out[1].TaktTimeModeZone_APLC_Out[1].Cycle_Done )
      wire#w5
      Contact( "Put Sinais de Interlock Falcare"."TURNO ATIVO FALCARE" )
      Coil( #barreira_invadida )
   END_RUNG
   RUNG wire#powerrail
      Contact( "Signals".ProcessInterlock_APLC_Input[1].ModezoneInterlock_APLC_Input[1].StationInterlock_APLC_Input[4].PositionInterlock_APLC_Input[1].EquipmentInterlock_APLC_Input[1].SignalInterlock_APLC_Input[7] )
   END_RUNG wire#w3
   RUNG wire#w4
      Contact( "AlwaysFALSE" )
      { S7_Templates := "SrcType := Time" } LT_Contact(in1 := "AREA_TaktTime.SIMPLE_INTERFACE_TAKTTIME_INPUT".TaktTimeWorkhop_APLC_Out[1].TaktTimeProcess_APLC_Out[1].TaktTimeModeZone_APLC_Out[1]."Timer", in2 := T#0s)
   END_RUNG wire#w5
   RUNG wire#powerrail
      Contact( #aciona_buzzer )
      wire#w6
      Coil( "Buzzer_P01" )
   END_RUNG
   RUNG wire#powerrail
      Contact( #barreira_invadida )
   END_RUNG wire#w6
   RUNG wire#w6
      Coil( "Buzzer_P40" )
   END_RUNG
   RUNG wire#powerrail
      Contact( #aciona_lampada_vermelha )
      wire#w7
      Coil( "Led_red_P01" )
   END_RUNG
   RUNG wire#powerrail
      Contact( #barreira_invadida )
   END_RUNG wire#w7
   RUNG wire#w7
      Coil( "Led_VermelhoP40" )
   END_RUNG
   RUNG wire#powerrail
      Contact( #aciona_lampada_verde )
      wire#w8
      Coil( "Led_verde_P01" )
   END_RUNG
   RUNG wire#w8
      Coil( "Led_VerdeP40" )
   END_RUNG
   // the same network as SCL:
   "Led_azul_P01" := "AREA_TaktTime.INTERFACE_TAKTTIME_INPUT".TaktTimeWorkhop_SPLC_Out[1].TaktTimeProcess_SPLC_Out[1].TaktTimeModeZone_SPLC_Out[2].StatusTakt = 2;
   "Led_azulP40" := "Led_azul_P01";
   "IEC_Timer_0_DB_20".TOF(IN := "AREA_TaktTime.SIMPLE_INTERFACE_TAKTTIME_INPUT".TaktTimeWorkhop_APLC_Out[1].TaktTimeProcess_APLC_Out[1].TaktTimeModeZone_APLC_Out[1]."Timer" = T#30s,
                           PT := T#5s);
   #aciona_buzzer := ("IEC_Timer_0_DB_20".Q AND "Clock_1.25Hz") OR ("Put Sinais de Interlock Falcare"."Moldezone 1 Done" AND NOT "IEC_Timer_0_DB_20".Q);
   #aciona_lampada_vermelha := #aciona_buzzer AND NOT "Put Sinais de Interlock Falcare"."Moldezone 1 Done";
   #aciona_lampada_verde := #aciona_buzzer;
   #barreira_invadida := ("Signals".ProcessInterlock_APLC_Input[1].ModezoneInterlock_APLC_Input[1].StationInterlock_APLC_Input[4].PositionInterlock_APLC_Input[1].EquipmentInterlock_APLC_Input[1].SignalInterlock_APLC_Input[6] OR "Signals".ProcessInterlock_APLC_Input[1].ModezoneInterlock_APLC_Input[1].StationInterlock_APLC_Input[4].PositionInterlock_APLC_Input[1].EquipmentInterlock_APLC_Input[1].SignalInterlock_APLC_Input[7]) AND ("AREA_TaktTime.SIMPLE_INTERFACE_TAKTTIME_INPUT".TaktTimeWorkhop_APLC_Out[1].TaktTimeProcess_APLC_Out[1].TaktTimeModeZone_APLC_Out[1]."Timer" <= T#5s) AND ("AREA_TaktTime.SIMPLE_INTERFACE_TAKTTIME_INPUT".TaktTimeWorkhop_APLC_Out[1].TaktTimeProcess_APLC_Out[1].TaktTimeModeZone_APLC_Out[1].Cycle_Done OR ("AlwaysFALSE" AND ("AREA_TaktTime.SIMPLE_INTERFACE_TAKTTIME_INPUT".TaktTimeWorkhop_APLC_Out[1].TaktTimeProcess_APLC_Out[1].TaktTimeModeZone_APLC_Out[1]."Timer" < T#0s))) AND "Put Sinais de Interlock Falcare"."TURNO ATIVO FALCARE";
   "Buzzer_P01" := #aciona_buzzer OR #barreira_invadida;
   "Buzzer_P40" := "Buzzer_P01";
   "Led_red_P01" := #aciona_lampada_vermelha OR #barreira_invadida;
   "Led_VermelhoP40" := "Led_red_P01";
   "Led_verde_P01" := #aciona_lampada_verde;
   "Led_VerdeP40" := #aciona_lampada_verde;
END_REGION

REGION Network 2 (SCL)
   IF "VERIFICA INTERLOCK"."ATIVA FOR" THEN
       FOR #INDEX_SIGNAL := 1 TO "Station_Setup_Const" DO
           FOR #INDEX_SIGNAL1 := 1 TO "Equipment_Setup_Const" DO
               FOR #INDEX_SIGNAL2 := 1 TO "Signal_Setup_Const" DO
                   IF "Signals".ProcessInterlock_APLC_Input[1].ModezoneInterlock_APLC_Input[2].StationInterlock_APLC_Input[#INDEX_SIGNAL]
                       .PositionInterlock_APLC_Input[1].EquipmentInterlock_APLC_Input[#INDEX_SIGNAL1].SignalInterlock_APLC_Input[#INDEX_SIGNAL2] = TRUE THEN
                       FOR #INDEX_VERIFICA := 1 TO 10 DO
                           IF "VERIFICA INTERLOCK".INTERLOCK[#INDEX_VERIFICA].STATION = 0 THEN
                               "VERIFICA INTERLOCK".INTERLOCK[#INDEX_VERIFICA].STATION := #INDEX_SIGNAL;
                               "VERIFICA INTERLOCK".INTERLOCK[#INDEX_VERIFICA].EQUIPAMENTO := #INDEX_SIGNAL1;
                               "VERIFICA INTERLOCK".INTERLOCK[#INDEX_VERIFICA].SINAL := #INDEX_SIGNAL2;
                               EXIT;
                           END_IF;
                       END_FOR;
                   END_IF;
                   END_FOR;
               END_FOR;
           END_FOR;
           "VERIFICA INTERLOCK"."ATIVA FOR" := FALSE;
       END_IF;
END_REGION

REGION Network 3
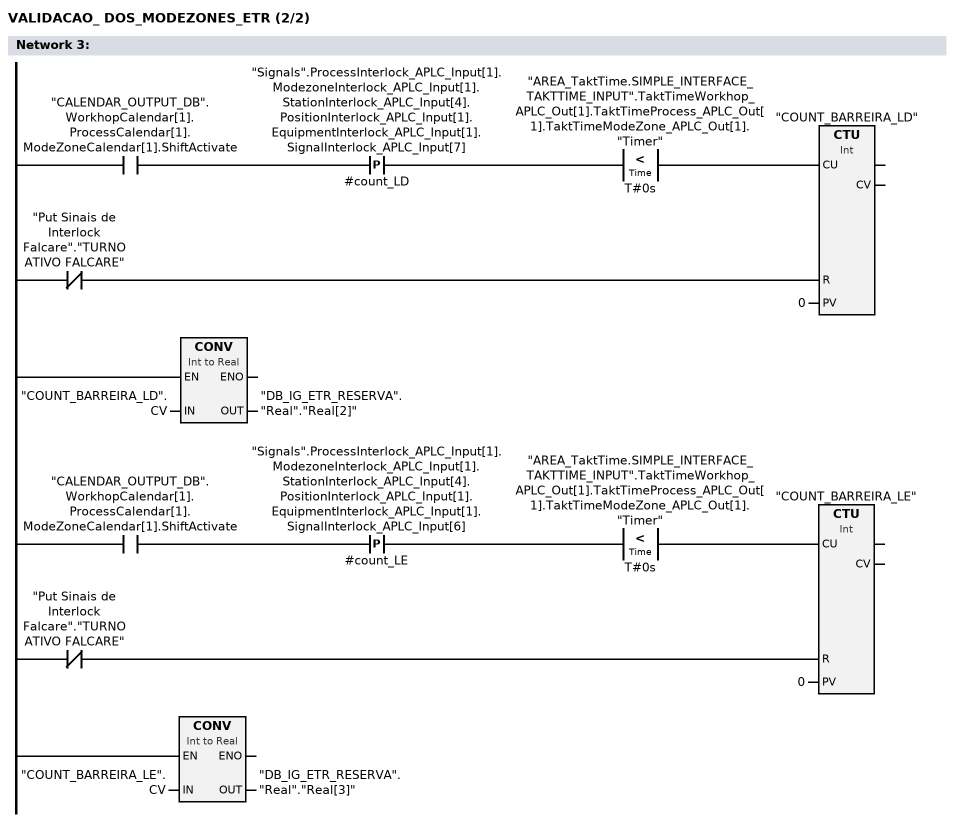
   RUNG wire#powerrail
      Contact( "CALENDAR_OUTPUT_DB".WorkhopCalendar[1].ProcessCalendar[1].ModeZoneCalendar[1].ShiftActivate )
      P_Contact(operand := "Signals".ProcessInterlock_APLC_Input[1].ModezoneInterlock_APLC_Input[1].StationInterlock_APLC_Input[4].PositionInterlock_APLC_Input[1].EquipmentInterlock_APLC_Input[1].SignalInterlock_APLC_Input[7], bit := #count_LD)
      { S7_Templates := "SrcType := Time" } LT_Contact(in1 := "AREA_TaktTime.SIMPLE_INTERFACE_TAKTTIME_INPUT".TaktTimeWorkhop_APLC_Out[1].TaktTimeProcess_APLC_Out[1].TaktTimeModeZone_APLC_Out[1]."Timer", in2 := T#0s)
      { S7_Templates := "value_type := Int" } "COUNT_BARREIRA_LD".CTU(r := wire#w1, pv := 0, cv =>)
   END_RUNG
   RUNG wire#powerrail
      I_Contact( "Put Sinais de Interlock Falcare"."TURNO ATIVO FALCARE" )
   END_RUNG wire#w1
   RUNG wire#powerrail
      { S7_Templates := "[SrcType := Int, DestType := Real]" } Convert(in := "COUNT_BARREIRA_LD".CV, out => "DB_IG_ETR_RESERVA"."Real"."Real[2]")
   END_RUNG
   RUNG wire#powerrail
      Contact( "CALENDAR_OUTPUT_DB".WorkhopCalendar[1].ProcessCalendar[1].ModeZoneCalendar[1].ShiftActivate )
      P_Contact(operand := "Signals".ProcessInterlock_APLC_Input[1].ModezoneInterlock_APLC_Input[1].StationInterlock_APLC_Input[4].PositionInterlock_APLC_Input[1].EquipmentInterlock_APLC_Input[1].SignalInterlock_APLC_Input[6], bit := #count_LE)
      { S7_Templates := "SrcType := Time" } LT_Contact(in1 := "AREA_TaktTime.SIMPLE_INTERFACE_TAKTTIME_INPUT".TaktTimeWorkhop_APLC_Out[1].TaktTimeProcess_APLC_Out[1].TaktTimeModeZone_APLC_Out[1]."Timer", in2 := T#0s)
      { S7_Templates := "value_type := Int" } "COUNT_BARREIRA_LE".CTU(r := wire#w2, pv := 0, cv =>)
   END_RUNG
   RUNG wire#powerrail
      I_Contact( "Put Sinais de Interlock Falcare"."TURNO ATIVO FALCARE" )
   END_RUNG wire#w2
   RUNG wire#powerrail
      { S7_Templates := "[SrcType := Int, DestType := Real]" } Convert(in := "COUNT_BARREIRA_LE".CV, out => "DB_IG_ETR_RESERVA"."Real"."Real[3]")
   END_RUNG
   // the same network as SCL:
   #_w1 := "CALENDAR_OUTPUT_DB".WorkhopCalendar[1].ProcessCalendar[1].ModeZoneCalendar[1].ShiftActivate AND "Signals".ProcessInterlock_APLC_Input[1].ModezoneInterlock_APLC_Input[1].StationInterlock_APLC_Input[4].PositionInterlock_APLC_Input[1].EquipmentInterlock_APLC_Input[1].SignalInterlock_APLC_Input[7] AND NOT #count_LD;   // rising edge of "Signals".ProcessInterlock_APLC_Input[1].ModezoneInterlock_APLC_Input[1].StationInterlock_APLC_Input[4].PositionInterlock_APLC_Input[1].EquipmentInterlock_APLC_Input[1].SignalInterlock_APLC_Input[7]
   #count_LD := "Signals".ProcessInterlock_APLC_Input[1].ModezoneInterlock_APLC_Input[1].StationInterlock_APLC_Input[4].PositionInterlock_APLC_Input[1].EquipmentInterlock_APLC_Input[1].SignalInterlock_APLC_Input[7];
   "COUNT_BARREIRA_LD".CTU(CU := #_w1 AND ("AREA_TaktTime.SIMPLE_INTERFACE_TAKTTIME_INPUT".TaktTimeWorkhop_APLC_Out[1].TaktTimeProcess_APLC_Out[1].TaktTimeModeZone_APLC_Out[1]."Timer" < T#0s),
                           R := NOT "Put Sinais de Interlock Falcare"."TURNO ATIVO FALCARE",
                           PV := 0);
   "DB_IG_ETR_RESERVA"."Real"."Real[2]" := INT_TO_REAL("COUNT_BARREIRA_LD".CV);
   #_w2 := "CALENDAR_OUTPUT_DB".WorkhopCalendar[1].ProcessCalendar[1].ModeZoneCalendar[1].ShiftActivate AND "Signals".ProcessInterlock_APLC_Input[1].ModezoneInterlock_APLC_Input[1].StationInterlock_APLC_Input[4].PositionInterlock_APLC_Input[1].EquipmentInterlock_APLC_Input[1].SignalInterlock_APLC_Input[6] AND NOT #count_LE;   // rising edge of "Signals".ProcessInterlock_APLC_Input[1].ModezoneInterlock_APLC_Input[1].StationInterlock_APLC_Input[4].PositionInterlock_APLC_Input[1].EquipmentInterlock_APLC_Input[1].SignalInterlock_APLC_Input[6]
   #count_LE := "Signals".ProcessInterlock_APLC_Input[1].ModezoneInterlock_APLC_Input[1].StationInterlock_APLC_Input[4].PositionInterlock_APLC_Input[1].EquipmentInterlock_APLC_Input[1].SignalInterlock_APLC_Input[6];
   "COUNT_BARREIRA_LE".CTU(CU := #_w2 AND ("AREA_TaktTime.SIMPLE_INTERFACE_TAKTTIME_INPUT".TaktTimeWorkhop_APLC_Out[1].TaktTimeProcess_APLC_Out[1].TaktTimeModeZone_APLC_Out[1]."Timer" < T#0s),
                           R := NOT "Put Sinais de Interlock Falcare"."TURNO ATIVO FALCARE",
                           PV := 0);
   "DB_IG_ETR_RESERVA"."Real"."Real[3]" := INT_TO_REAL("COUNT_BARREIRA_LE".CV);
END_REGION
END_FUNCTION

FUNCTION "ALARMES" : Void   // FC13, LAD
{ S7_Optimized_Access := 'TRUE' }
// stored: SetENOAutomatically false
BEGIN

REGION Network 1: ALARMES CABINE
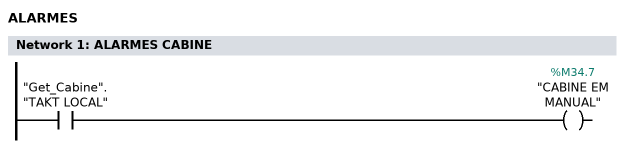
   RUNG wire#powerrail
      Contact( "Get_Cabine"."TAKT LOCAL" )
      Coil( "CABINE EM MANUAL" )
   END_RUNG
   // the same network as SCL:
   "CABINE EM MANUAL" := "Get_Cabine"."TAKT LOCAL";
END_REGION
END_FUNCTION

FUNCTION "Clock" : Void
{ S7_Optimized_Access := 'TRUE' }
VERSION : 0.1
   VAR_TEMP 
      ret : Int;
   END_VAR


BEGIN
	#ret := RD_LOC_T("General_functions".Clock.DateTime);
END_FUNCTION

ORGANIZATION_BLOCK "Programming error"

{ S7_Optimized_Access := 'TRUE' }
VERSION : 0.1
VAR_INPUT
  BlockNr : UInt;(*Number of causing block*)
  Reaction : USInt;(*0:ignore, 1:substitute, 2:skip*)
  Fault_ID : Byte;(*Fault identifier*)
  BlockType : USInt;(*16#01:OB, 16#02:FC, 16#03:FB, 16#04:SFC, 16#05:SFB, 16#06:DB: Type of block causing the error*)
  Area : USInt;(*Area where the error occured*)
  DBNr : DB_ANY;(*DB number if Area = DB or DI*)
  Csg_OBNr : OB_ANY;(*Number of OB causing the error*)
  Csg_Prio : USInt;(*Priority of OB causing the error*)
  Width : USInt;(*0:bit, 1:byte, 2:word, 3:dword, 4:lword*)
END_VAR

VAR_TEMP

END_VAR

VAR CONSTANT

END_VAR




BEGIN
END_ORGANIZATION_BLOCK
